   VAR CONSTANT
      C_REF_FREQUENCY : Int := 6000;   // [rpm]
      C_REF_VOLTAGE : Int := 1000;   // [V]
      C_REF_CURRENT : Int := 10;   // [A]
      C_REF_TORQUE : Int := 100;   // [Nm]
      C_REF_POWER : Int := 31;   // [W]
      C_REF_TEMP : Int := 100;   // [°C]
   END_VAR


BEGIN
	REGION Telegram Module
	    #t_ZSW1_Word := 0;
	    #t_POS_ZSW1_Word := 0;
	    #t_POS_ZSW2_Word := 0;
	    #t_ZSW2_Word := 0;

	    #t_Ret_Val_Int := RD_ADDR(LADDR := #i_Telegram_HW_ID,
	                              PIADDR => #t_HW_RD_Inf_Rec_I_Address,
	                              PICount => #t_HW_RD_Inf_Rec_I_Len,
	                              PQADDR => #t_HW_WR_Inf_Rec_O_Address,
	                              PQCount => #t_HW_WR_Inf_Rec_O_Len);

	    #o_Telegram_Start_Address := UDINT_TO_INT(#t_HW_RD_Inf_Rec_I_Address);

	    IF #t_Ret_Val_Int = 0 AND #t_HW_RD_Inf_Rec_I_Len = 24 THEN
	        // PZD1: ZSW1 (Word)
	        #t_ZSW1_Word := PEEK_WORD(area := 16#81, // Input area
	                                  dbNumber := 0,
	                                  byteOffset := UDINT_TO_DINT(#t_HW_RD_Inf_Rec_I_Address));

	        // PZD2: POS_ZSW1 (Word)
	        #t_POS_ZSW1_Word := PEEK_WORD(area := 16#81,
	                                      dbNumber := 0,
	                                      byteOffset := UDINT_TO_DINT(#t_HW_RD_Inf_Rec_I_Address) + 2);

	        // PZD3: POS_ZSW2 (Word)
	        #t_POS_ZSW2_Word := PEEK_WORD(area := 16#81,
	                                      dbNumber := 0,
	                                      byteOffset := UDINT_TO_DINT(#t_HW_RD_Inf_Rec_I_Address) + 4);

	        // PZD4: ZSW2 (Word)
	        #t_ZSW2_Word := PEEK_WORD(area := 16#81,
	                                  dbNumber := 0,
	                                  byteOffset := UDINT_TO_DINT(#t_HW_RD_Inf_Rec_I_Address) + 6);

	        // PZD5: Reserved (Int)
	        #o_Data.Reserved := 0;

	        // PZD6-7: XIST (Real/Float32) - Position actual value
	        #o_Data.XIST := DWORD_TO_REAL(PEEK_DWORD(area := 16#81,
	                                                                               dbNumber := 0,
	                                                                               byteOffset := UDINT_TO_DINT(#t_HW_RD_Inf_Rec_I_Address) + 10));

	        // PZD8-9: VIST (Real/Float32) - Velocity actual value
	        #o_Data.VIST := DWORD_TO_REAL(PEEK_DWORD(area := 16#81,
	                                                                               dbNumber := 0,
	                                                                               byteOffset := UDINT_TO_DINT(#t_HW_RD_Inf_Rec_I_Address) + 14));

	        // PZD10: MELDW (Word)
	        #o_Data.MELDW_Bit00_PositioningAbsolute := FALSE; // MELDW reserved in telegram 112

	        // PZD11: FaultCode (Word)
	        #o_Data.FaultCode := PEEK_WORD(area := 16#81,
	                                       dbNumber := 0,
	                                       byteOffset := UDINT_TO_DINT(#t_HW_RD_Inf_Rec_I_Address) + 20);

	        // PZD12: AlarmCode (Word)
	        #o_Data.AlarmCode := PEEK_WORD(area := 16#81,
	                                      dbNumber := 0,
	                                      byteOffset := UDINT_TO_DINT(#t_HW_RD_Inf_Rec_I_Address) + 22);
	    ELSE
	        #o_Data.XIST := 0.0;
	        #o_Data.VIST := 0.0;
	        #o_Data.FaultCode := 0;
	        #o_Data.AlarmCode := 0;
	    END_IF;

	    // Unpack ZSW1 bits
	    #o_Data.ZSW1_Bit00_ReadyOn := #t_ZSW1_Word.%X0;
	    #o_Data.ZSW1_Bit01_Ready := #t_ZSW1_Word.%X1;
	    #o_Data.ZSW1_Bit02_Enabled := #t_ZSW1_Word.%X2;
	    #o_Data.ZSW1_Bit03_Fault := #t_ZSW1_Word.%X3;
	    #o_Data.ZSW1_Bit04_Off2Inactive := #t_ZSW1_Word.%X4;
	    #o_Data.ZSW1_Bit05_Off3Inactive := #t_ZSW1_Word.%X5;
	    #o_Data.ZSW1_Bit06_Inhibit := #t_ZSW1_Word.%X6;
	    #o_Data.ZSW1_Bit07_Alarm := #t_ZSW1_Word.%X7;
	    #o_Data.ZSW1_Bit08_FollowingOK := #t_ZSW1_Word.%X8;
	    #o_Data.ZSW1_Bit09_Control := #t_ZSW1_Word.%X9;
	    #o_Data.ZSW1_Bit10_TargetReached := #t_ZSW1_Word.%X10;
	    #o_Data.ZSW1_Bit11_HomeSet := #t_ZSW1_Word.%X11;
	    #o_Data.ZSW1_Bit12_AckActive := #t_ZSW1_Word.%X12;
	    #o_Data.ZSW1_Bit13_SetpointFixed := #t_ZSW1_Word.%X13;
	    #o_Data.ZSW1_Bit14_AxisAccel := #t_ZSW1_Word.%X14;
	    #o_Data.ZSW1_Bit15_AxisDecel := #t_ZSW1_Word.%X15;

	    // Unpack POS_ZSW1 bits
	    #o_Data.POS_ZSW1_Bit00_Active0 := #t_POS_ZSW1_Word.%X0;
	    #o_Data.POS_ZSW1_Bit01_Active1 := #t_POS_ZSW1_Word.%X1;
	    #o_Data.POS_ZSW1_Bit02_Active2 := #t_POS_ZSW1_Word.%X2;
	    #o_Data.POS_ZSW1_Bit03_Active3 := #t_POS_ZSW1_Word.%X3;
	    #o_Data.POS_ZSW1_Bit04_Active4 := #t_POS_ZSW1_Word.%X4;
	    #o_Data.POS_ZSW1_Bit05_Active5 := #t_POS_ZSW1_Word.%X5;
	    #o_Data.POS_ZSW1_Bit06_Reserved := #t_POS_ZSW1_Word.%X6;
	    #o_Data.POS_ZSW1_Bit07_ReleaseBrake := #t_POS_ZSW1_Word.%X7;
	    #o_Data.POS_ZSW1_Bit08_StopCamMinus := #t_POS_ZSW1_Word.%X8;
	    #o_Data.POS_ZSW1_Bit09_StopCamPlus := #t_POS_ZSW1_Word.%X9;
	    #o_Data.POS_ZSW1_Bit10_JogActive := #t_POS_ZSW1_Word.%X10;
	    #o_Data.POS_ZSW1_Bit11_RefApproach := #t_POS_ZSW1_Word.%X11;
	    #o_Data.POS_ZSW1_Bit12_FlyingHoming := #t_POS_ZSW1_Word.%X12;
	    #o_Data.POS_ZSW1_Bit13_Traversing := #t_POS_ZSW1_Word.%X13;
	    #o_Data.POS_ZSW1_Bit14_Setup := #t_POS_ZSW1_Word.%X14;
	    #o_Data.POS_ZSW1_Bit15_MDI := #t_POS_ZSW1_Word.%X15;

	    // Unpack POS_ZSW2 bits
	    #o_Data.POS_ZSW2_Bit00_Tracking := #t_POS_ZSW2_Word.%X0;
	    #o_Data.POS_ZSW2_Bit01_VelLimit := #t_POS_ZSW2_Word.%X1;
	    #o_Data.POS_ZSW2_Bit02_TargetReached := #t_POS_ZSW2_Word.%X2;
	    #o_Data.POS_ZSW2_Bit03_PrintMark := #t_POS_ZSW2_Word.%X3;
	    #o_Data.POS_ZSW2_Bit04_Forward := #t_POS_ZSW2_Word.%X4;
	    #o_Data.POS_ZSW2_Bit05_Backward := #t_POS_ZSW2_Word.%X5;
	    #o_Data.POS_ZSW2_Bit06_SWLimitMinus := #t_POS_ZSW2_Word.%X6;
	    #o_Data.POS_ZSW2_Bit07_SWLimitPlus := #t_POS_ZSW2_Word.%X7;
	    #o_Data.POS_ZSW2_Bit08_Cam1 := #t_POS_ZSW2_Word.%X8;
	    #o_Data.POS_ZSW2_Bit09_Cam2 := #t_POS_ZSW2_Word.%X9;
	    #o_Data.POS_ZSW2_Bit10_Output1 := #t_POS_ZSW2_Word.%X10;
	    #o_Data.POS_ZSW2_Bit11_Output2 := #t_POS_ZSW2_Word.%X11;
	    #o_Data.POS_ZSW2_Bit12_FixedStop := #t_POS_ZSW2_Word.%X12;
	    #o_Data.POS_ZSW2_Bit13_Clamping := #t_POS_ZSW2_Word.%X13;
	    #o_Data.POS_ZSW2_Bit14_TravelFixed := #t_POS_ZSW2_Word.%X14;
	    #o_Data.POS_ZSW2_Bit15_TraversingCmd := #t_POS_ZSW2_Word.%X15;

	    // Unpack ZSW2 bits
	    #o_Data.ZSW2_Bit00_Reserved := #t_ZSW2_Word.%X0;
	    #o_Data.ZSW2_Bit01_Reserved := #t_ZSW2_Word.%X1;
	    #o_Data.ZSW2_Bit02_Reserved := #t_ZSW2_Word.%X2;
	    #o_Data.ZSW2_Bit03_Reserved := #t_ZSW2_Word.%X3;
	    #o_Data.ZSW2_Bit04_Reserved := #t_ZSW2_Word.%X4;
	    #o_Data.ZSW2_Bit05_Reserved := #t_ZSW2_Word.%X5;
	    #o_Data.ZSW2_Bit06_Reserved := #t_ZSW2_Word.%X6;
	    #o_Data.ZSW2_Bit07_Reserved := #t_ZSW2_Word.%X7;
	    #o_Data.ZSW2_Bit08_Reserved := #t_ZSW2_Word.%X8;
	    #o_Data.ZSW2_Bit09_Reserved := #t_ZSW2_Word.%X9;
	    #o_Data.ZSW2_Bit10_Reserved := #t_ZSW2_Word.%X10;
	    #o_Data.ZSW2_Bit11_Reserved := #t_ZSW2_Word.%X11;
	    #o_Data.ZSW2_Bit12_Reserved := #t_ZSW2_Word.%X12;
	    #o_Data.ZSW2_Bit13_Reserved := #t_ZSW2_Word.%X13;
	    #o_Data.ZSW2_Bit14_Reserved := #t_ZSW2_Word.%X14;
	    #o_Data.ZSW2_Bit15_Reserved := #t_ZSW2_Word.%X15;
	END_REGION

	REGION Actual Value Module (Extended Data)
	    #t_ZSW_S210_Word := 0;

	    #t_Ret_Val_Int := RD_ADDR(LADDR := #i_Additional_HW_ID,
	                              PIADDR => #t_HW_RD_Inf_Rec_I_Address,
	                              PICount => #t_HW_RD_Inf_Rec_I_Len,
	                              PQADDR => #t_HW_WR_Inf_Rec_O_Address,
	                              PQCount => #t_HW_WR_Inf_Rec_O_Len);

	    #o_ActualValue_Start_Address := UDINT_TO_INT(#t_HW_RD_Inf_Rec_I_Address);

	    IF #t_Ret_Val_Int = 0 AND #t_HW_RD_Inf_Rec_I_Len = 12 THEN
	        // Read ZSW_S210 (DI status word)
	        #t_ZSW_S210_Word := PEEK_WORD(area := 16#81, // Input area
	                                      dbNumber := 0,
	                                      byteOffset := UDINT_TO_DINT(#t_HW_RD_Inf_Rec_I_Address));

	        // Read DC Link Voltage (Int)
	        #t_Word_Scale_Data := PEEK_WORD(area := 16#81,
	                                        dbNumber := 0,
	                                        byteOffset := UDINT_TO_DINT(#t_HW_RD_Inf_Rec_I_Address) + 2);

	        #o_Data.DCLinkVoltage := DINT_TO_INT(WORD_TO_DINT(#t_Word_Scale_Data) * #C_REF_VOLTAGE / 16#4000);

	        // Read Actual Current (Int)
	        #t_Word_Scale_Data := PEEK_WORD(area := 16#81,
	                                        dbNumber := 0,
	                                        byteOffset := UDINT_TO_DINT(#t_HW_RD_Inf_Rec_I_Address) + 4);

	        #o_Data.ActualCurrent := DINT_TO_INT(WORD_TO_DINT(#t_Word_Scale_Data) * #C_REF_CURRENT * 10 / 16#4000);

	        // Read Active Power (Int)
	        #t_Word_Scale_Data := PEEK_WORD(area := 16#81,
	                                        dbNumber := 0,
	                                        byteOffset := UDINT_TO_DINT(#t_HW_RD_Inf_Rec_I_Address) + 6);

	        #o_Data.ActivePower := DINT_TO_INT(WORD_TO_DINT(#t_Word_Scale_Data) * #C_REF_POWER / 16#4000);

	        // Read Active Utilization (Int)
	        #t_Word_Scale_Data := PEEK_WORD(area := 16#81,
	                                        dbNumber := 0,
	                                        byteOffset := UDINT_TO_DINT(#t_HW_RD_Inf_Rec_I_Address) + 8);

	        #o_Data.TorqueUtilization := DINT_TO_INT(WORD_TO_DINT(#t_Word_Scale_Data) * 100 / 16#4000);

	        // Read Motor Load Rate (Int)
	        #t_Word_Scale_Data := PEEK_WORD(area := 16#81,
	                                        dbNumber := 0,
	                                        byteOffset := UDINT_TO_DINT(#t_HW_RD_Inf_Rec_I_Address) + 10);

	        #o_Data.MotorUtilization := DINT_TO_INT(WORD_TO_DINT(#t_Word_Scale_Data) * 100 / 16#4000);
	    ELSE
	        #o_Data.DCLinkVoltage := 0;
	        #o_Data.ActualCurrent := 0;
	        #o_Data.ActivePower := 0;
	        #o_Data.TorqueUtilization := 0;
	        #o_Data.MotorUtilization := 0;
	    END_IF;

	    // Unpack ZSW_S210 bits (DI status)
	    #o_Data.ZSW_S210_Bit00_DI0 := #t_ZSW_S210_Word.%X0;
	    #o_Data.ZSW_S210_Bit01_DI1 := #t_ZSW_S210_Word.%X1;
	    #o_Data.ZSW_S210_Bit02_DI2 := #t_ZSW_S210_Word.%X2;
	    #o_Data.ZSW_S210_Bit03_DI3 := #t_ZSW_S210_Word.%X3;
	    #o_Data.ZSW_S210_Bit04_DI4 := #t_ZSW_S210_Word.%X4;
	    #o_Data.ZSW_S210_Bit05_Reserved := #t_ZSW_S210_Word.%X5;
	    #o_Data.ZSW_S210_Bit06_Reserved := #t_ZSW_S210_Word.%X6;
	    #o_Data.ZSW_S210_Bit07_Reserved := #t_ZSW_S210_Word.%X7;
	    #o_Data.ZSW_S210_Bit08_Reserved := #t_ZSW_S210_Word.%X8;
	    #o_Data.ZSW_S210_Bit09_Reserved := #t_ZSW_S210_Word.%X9;
	    #o_Data.ZSW_S210_Bit10_Reserved := #t_ZSW_S210_Word.%X10;
	    #o_Data.ZSW_S210_Bit11_Reserved := #t_ZSW_S210_Word.%X11;
	    #o_Data.ZSW_S210_Bit12_Reserved := #t_ZSW_S210_Word.%X12;
	    #o_Data.ZSW_S210_Bit13_Reserved := #t_ZSW_S210_Word.%X13;
	    #o_Data.ZSW_S210_Bit14_Reserved := #t_ZSW_S210_Word.%X14;
	    #o_Data.ZSW_S210_Bit15_Reserved := #t_ZSW_S210_Word.%X15;
	END_REGION
END_FUNCTION

TYPE "UDT_S210_SW_Output"
VERSION : 0.1
   STRUCT
      AxisEnabled : Bool;   // 驱动已使能
      AxisPosOk : Bool;   // 目标位置到达
      AxisSpFixed : Bool;   // 设定位置到达
      AxisRef : Bool;   // 已设置参考点
      AxisWarn : Bool;   // 驱动报警
      AxisError : Bool;   // 驱动故障
      Lockout : Bool;   // 禁止接通
      ActVelocity : Real;   // 实际速度
      ActPosition : Real;   // 当前位置
      ActMode : Int;   // 当前激活的运行模式
      EPosZSW1 : Word;   // POS ZSW1的状态
      EPosZSW2 : Word;   // POS ZSW2的状态
      AlarmCode : Word;   // 驱动器当前的报警代码
      FaultCode : Word;   // 驱动器当前的故障代码
      ZSW1 : Word;   // ZSW1的状态
      ZSW2 : Word;   // ZSW2的状态
      MELDW : Word;   // MELDW的状态
      Error : Bool;   // 1=存在错误
      Status : Word;   // 16#7002：无故障，正常运行
      DiagID : Word;   // 扩展的通信错误
   END_STRUCT;

END_TYPE

TYPE "UDT_S210_SW_Input"
VERSION : 0.1
   STRUCT
      Mode : Int;
      Enbale : Bool;
      CancelTraversing : Bool;
      IntermediateStop : Bool;
      Positive : Bool;
      Negative : Bool;
      Jog_Left : Bool;
      Jog_Right : Bool;
      FlyRef : Bool;
      AckError : Bool;
      ExecuteMode : Bool;
      Position : Real;
      Velocity : Real;
      OverV : Int;
      Acceleration : Real;
      Deceleration : Real;
      FixStopTorque : Real;
      RefCoordinate : Real;
      ConfigEPOS : DWord;
   END_STRUCT;

END_TYPE

FUNCTION_BLOCK "FB_SINA_POS_TEL112"
{ S7_Optimized_Access := 'TRUE' }
VERSION : 0.2
   VAR_INPUT
      modePos : Int;   // Settings of the mode
      enableAxis : Bool;   // 1 = Enable the drive
      cancelTraversing : Bool := TRUE;   // 0 = Reject active traverse task
      intermediateStop : Bool := TRUE;   // 0 = Intermediate STOP of traverse command
      positive : Bool;   // 1 = Direction positive
      negative : Bool;   // 1 = Direction negative
      jog1 : Bool;   // 1 = Use jog 1 (direction / speed)
      jog2 : Bool;   // 1 = Use jog 2 (direction / speed)
      flyRef : Bool;   // 1 = Start flying reference function
      ackError : Bool;   // 1  = Acknowledge of errors
      executeMode : Bool;   // 0-->1 = Start the mode
      position : Real;   // Position of the MDI mode or setting of traversing block
      velocity : Real;   // MDI velocity
      overV : Int := 100;   // Override of  velocity in [%] --> 4000h=100%
      acceleration : Real;   // MDI acceleration
      deceleration : Real;   // MDI deceleration
      fixStopTorque : Real;   // torque setting for fix stop function (reserved)
      refCoordinate : Real;
      configEPOS : DWord := 16#0000_0003;   // binary programmed input to control all functions in the telegram without its own function block input
   END_VAR

   VAR_OUTPUT
      axisEnabled : Bool;   // 1= Axis in operation
      axisPosOk : Bool;   // 1= Position setpoint reached
      axisSpFixed : Bool;   // 1= Setpoint fixed (Attention: Dependence on SINAMICS firmware)
      axisRef : Bool;   // 1= Reference point set
      axisWarn : Bool;   // 1= Axis alarm / warning present
      axisError : Bool;   // 1= Axis fault present
      lockOut : Bool;   // 1= Axis in lockout state
      actVelocity : Real;   // actual axis velocity
      actPosition : Real;   // actual axis position
      actMode : Int;   // Active EPos mode
      actWarn : Word;   // Actual number of warning
      actFault : Word;   // Actual number of error
      error : Bool;   // 1 = Error  (FB and Infeed)
      status : Word;   // Status output (7002 = FB in operation; 8xxx = error description  - read the manual)
      diagID : Word;   // Error codes of the cyclic system funtion blocks DPWR / DPRD_DAT (固定为0)
   END_VAR

   VAR_IN_OUT
      InputData : "UDT_S210_HW_Input";   // 从驱动器接收的数据
      OutputData : "UDT_S210_HW_Output";   // 发送到驱动器的数据
   END_VAR

   VAR
      sbOff1Edge : Bool := 0;   // Positive edge of starting or stopping the device
      sbOff1 : Bool := 0;   // Starting or stopping the device
      sbExecuteEdge : Bool := 0;   // Positive edge of activate traversing block
      sbExecute : Bool := 0;   // Activate traversing block
      sbRefTypEdge : Bool := 0;   // Positive edge of referencing type "flying reference"
      sbRefTyp : Bool := 0;   // Referencing type "flying reference"
      sbMdiStart : Bool := 0;   // Direct setpoint input / MDI - start
      sbMdiStartEdge : Bool := 0;   // Positive edge of direct setpoint input / MDI - start
      sbRefStart : Bool := 0;   // Referencing start
      sbJogInc : Bool := 0;   // Jogging incremental
      sbReady : Bool := 0;   // Ready to power up / to start
      sbIOp : Bool := 0;   // Ready to operate
      sbAccel : Bool := 0;   // Axis accelerating
      sbDecel : Bool := 0;   // Axis decelerating
      sbAlarm : Bool := 0;   // Alarm / Warnung present
      sbFault : Bool := 0;   // Fault present
      sbFWD : Bool := 0;   // Axis drives forwards
      sbBWD : Bool := 0;   // Axis drives backwards
      sbBusy : Bool := 0;   // Mode of operation is explained
      swStatus : Word := 16#0000;   // Mode of operation disturbance
      siExecuteCyc : Int := 0;   // Counter of runcycle of active traversing block
      siRefTypCyc : Int := 0;   // Counter of runcycle of referencing type "flying reference"
      siJogIncCyc : Int := 0;   // Counter of runcycle of jogging incremental
      siMdiStartCyc : Int := 0;   // Counter of runcycle of direct setpoint input / MDI - start
      siRefActRetry : Int := 0;   // Counter of retry of reference point approach active
      siModePos : Int := 0;   // Setting of mode
      siCycWait : Int := 5;   // Counter of cycle of waiting
      siRetryMax : Int := 30;   // Max. count of cycles of retry
      sbModePos : Bool := 0;   // Mode of setting okay
   END_VAR

   VAR CONSTANT
      MODEPOSMAX : Int := 9;   // Max. count of mode
      TRAVERSEBLOCKMAXNO : Int := 32;   // Max. number of traversing block
   END_VAR


BEGIN
	//=============================================================================
	//SIEMENS AG
	//(c)Copyright 2023 All Rights Reserved
	//-----------------------------------------------------------------------------
	// Library: DriveLib
	// Tested with: -
	// Engineering: TIA Portal V18
	// Restrictions: -
	// Requirements: S7-1200 / S7-1500
	// Functionality: cyclic communication between a SINAMICS (Basic positioner)and a PLC
	//                If in HWConfig Std.TLG 112 is projected 17/12 PZD-words are exchanged
	//                in every bus cycle.
	//                The parametrisation of these words is described in the manual of the
	//                SINAMICS
	// Contactor: mc_gmc_mp_asia.cn@siemens.com
	// *****************************************************************************
	// Version:
	// V0.0: Created
	// V0.2: 重构 - 移除DPWR/DPRD，改用外部UDT (UDT_S210_HW_Output/Input)
	//=============================================================================

	// The input of the modePos should between 1 and the MODEPOSMAX
	IF #modePos > #MODEPOSMAX OR #modePos < 1 THEN
	    #sbModePos := FALSE;
	    #error := True;
	    #swStatus := 16#8202;
	ELSE
	    IF NOT #sbFWD AND NOT #sbBWD AND NOT #sbAccel AND NOT #sbDecel THEN
	        #sbModePos := TRUE;
	        #siModePos := #modePos;
	        IF #swStatus = 16#8202 THEN
	            #swStatus := 16#7002;
	            #error := False;
	        END_IF;
	    END_IF;
	END_IF;

	// Check the overrider setting
	IF (#overV < 0) OR (#overV > 199) THEN
	    #swStatus := 16#8203;
	    #error := True;
	ELSE
	    // Override映射到OutputData.Override (Int类型，0-16384对应0-100%)
	    #OutputData.Override := REAL_TO_INT(16384.0 * (INT_TO_REAL(#overV) / 100.0));
	END_IF;

	// Check the acceleration and deceleration setting
	IF #acceleration < 0.0 THEN
	    #swStatus := 16#8203;
	    #error := True;
	ELSE
	    #OutputData.MDI_ACC := #acceleration;
	END_IF;
	IF #deceleration < 0.0 THEN
	    #swStatus := 16#8203;
	    #error := True;
	ELSE
	    #OutputData.MDI_DEC := #deceleration;
	END_IF;
	IF NOT (#overV < 0) AND NOT (#overV > 199) AND NOT (#acceleration < 0.0) AND NOT (#deceleration < 0.0) THEN
	    IF #swStatus = 16#8203 THEN
	        #swStatus := 16#7002;
	        #error := FALSE;
	    END_IF;
	END_IF;

	// 位置、速度、参考坐标直接映射
	#OutputData.MDI_TARPOS := #position;
	#OutputData.MDI_VELOCITY := #velocity;
	#OutputData.REF_COORDINATE := #refCoordinate;

	// Enable the axis
	IF #enableAxis AND NOT #sbOff1Edge AND NOT #sbBusy AND #sbModePos THEN
	    #sbOff1 := True;
	END_IF;
	#sbOff1Edge := #enableAxis AND NOT #sbBusy;
	IF NOT #enableAxis THEN
	    #sbOff1 := False;
	END_IF;

	// Flying reference
	IF #flyRef AND NOT #sbRefTypEdge THEN
	    #sbRefTyp := True;
	END_IF;
	#sbRefTypEdge := #flyRef;
	IF NOT #flyRef THEN
	    #sbRefTyp := False;
	    #siRefTypCyc := 0;
	END_IF;

	// Execute the motion
	IF #executeMode AND NOT #sbExecuteEdge THEN
	    #sbExecute := True;
	    #siExecuteCyc := 0;
	ELSIF #actMode <> #modePos THEN
	    #sbExecute := FALSE;
	ELSIF #siExecuteCyc > (15 * #siCycWait) THEN
	    IF #modePos <> 4 THEN
	        #sbExecute := FALSE;
	    ELSE
	        // 使用InputData.ZSW1_Bit11_HomeSet替代sxRecvBuf.ZSW1.%X11
	        IF #InputData.ZSW1_Bit11_HomeSet OR NOT #executeMode THEN
	            #sbExecute := FALSE;
	        END_IF;
	    END_IF;
	ELSE
	    ;
	END_IF;
	IF #siExecuteCyc > 100 THEN
	    #siExecuteCyc := 0;
	ELSE
	    #siExecuteCyc := #siExecuteCyc + 1;
	END_IF;
	#sbExecuteEdge := #executeMode;

	// MDI Start边沿检测逻辑（基于EPosSTW1.%X15，即POS_STW1_Bit15_ActivateMDI）
	IF #OutputData.POS_STW1_Bit15_ActivateMDI AND NOT #sbMdiStartEdge THEN
	    #sbMdiStart := True;
	END_IF;
	#sbMdiStartEdge := #OutputData.POS_STW1_Bit15_ActivateMDI AND NOT #sbBusy;
	IF NOT #OutputData.POS_STW1_Bit15_ActivateMDI THEN
	    #sbMdiStart := False;
	    #siMdiStartCyc := 0;
	END_IF;

	// 基础STW1控制位映射
	#OutputData.STW1_Bit04_NotRejectTask := #cancelTraversing;
	#OutputData.STW1_Bit05_NoIntermediateStop := #intermediateStop;
	#OutputData.STW1_Bit07_Ack := #ackError;
	#OutputData.STW1_Bit01_Off2 := TRUE;  // 原.%X1
	#OutputData.STW1_Bit02_Off3 := TRUE;  // 原.%X2
	#OutputData.STW1_Bit03_Enable := TRUE; // 原.%X3
	#OutputData.STW1_Bit10_PLC := TRUE;    // 原.%X10 (Life bit)
	#OutputData.STW1_Bit12_Reserved := FALSE; // 原.%X12
	#OutputData.STW1_Bit14_Reserved := FALSE; // 原.%X14
	#OutputData.STW1_Bit15_Reserved := FALSE; // 原.%X15

	// If the parameter setting is correnct, then execute the positioning mode.
	// ModePos = 1, relative positioning
	IF (#siModePos = 1 AND #sbModePos) THEN
	    #OutputData.STW1_Bit00_On := #sbOff1;           // 原STW1.%X0
	    #OutputData.STW1_Bit08_Jog1 := False;           // 原.%X8
	    #OutputData.STW1_Bit09_Jog2 := False;           // 原.%X9
	    #OutputData.STW1_Bit11_StartHoming := False;    // 原.%X11

	    #OutputData.POS_STW1_Bit08_Absolute := False;    // 原EPosSTW1.%X8 (0=相对)
	    #OutputData.POS_STW1_Bit09_DirPos := False;      // 原.%X9
	    #OutputData.POS_STW1_Bit10_DirNeg := False;      // 原.%X10
	    #OutputData.POS_STW1_Bit14_SetupOrPositioning := False; // 原.%X14 (0=定位)
	    #OutputData.POS_STW1_Bit15_ActivateMDI := False; // 原.%X15

	    #OutputData.POS_STW2_Bit01_SetRefPoint := False;  // 原.%X1
	    #OutputData.POS_STW2_Bit03_AdjustEncoder := False; // 原.%X3
	    #OutputData.POS_STW2_Bit05_JogIncrementalOrVelocity := False; // 原.%X5
	    #OutputData.POS_STW2_Bit09_RefNegDir := False;    // 原.%X9
	    #OutputData.POS_STW2_Bit08_RefType := False;      // 原.%X8

	    IF #sbOff1 AND #sbReady AND #sbIOp AND NOT #sbFault THEN
	        #OutputData.POS_STW1_Bit15_ActivateMDI := True;  // MDI激活
	        #OutputData.POS_STW1_Bit08_Absolute := False;    // 相对定位
	        IF #positive AND NOT #negative THEN
	            #OutputData.POS_STW1_Bit09_DirPos := True;
	            #OutputData.POS_STW1_Bit10_DirNeg := False;
	        ELSIF NOT #positive AND #negative THEN
	            #OutputData.POS_STW1_Bit09_DirPos := False;
	            #OutputData.POS_STW1_Bit10_DirNeg := True;
	        ELSE
	            #OutputData.POS_STW1_Bit09_DirPos := False;
	            #OutputData.POS_STW1_Bit10_DirNeg := False;
	        END_IF;
	        IF #sbMdiStart AND (#siMdiStartCyc < #siCycWait) THEN
	            #siMdiStartCyc := #siMdiStartCyc + 1;
	        ELSE
	            #OutputData.STW1_Bit06_ActivateTask := #sbExecute; // 原.%X6
	        END_IF;
	        IF #sbRefTyp THEN
	            #OutputData.POS_STW2_Bit08_RefType := True; // 飞参模式
	            IF (#siRefTypCyc = 0) THEN
	                #siRefTypCyc := #siRefTypCyc + 1;
	            ELSE
	                #OutputData.STW1_Bit11_StartHoming := True; // 开始回零
	            END_IF;
	        END_IF;
	    END_IF;

	    // ModePos = 2, absolute positioning
	ELSIF (#siModePos = 2 AND #sbModePos) THEN
	    #OutputData.STW1_Bit00_On := #sbOff1;
	    #OutputData.STW1_Bit08_Jog1 := False;
	    #OutputData.STW1_Bit09_Jog2 := False;
	    #OutputData.STW1_Bit11_StartHoming := False;

	    #OutputData.POS_STW1_Bit08_Absolute := False;
	    #OutputData.POS_STW1_Bit09_DirPos := False;
	    #OutputData.POS_STW1_Bit10_DirNeg := False;
	    #OutputData.POS_STW1_Bit14_SetupOrPositioning := False;
	    #OutputData.POS_STW1_Bit15_ActivateMDI := False;

	    #OutputData.POS_STW2_Bit01_SetRefPoint := False;
	    #OutputData.POS_STW2_Bit03_AdjustEncoder := False;
	    #OutputData.POS_STW2_Bit05_JogIncrementalOrVelocity := False;
	    #OutputData.POS_STW2_Bit09_RefNegDir := False;
	    #OutputData.POS_STW2_Bit08_RefType := False;

	    IF #sbOff1 AND #sbReady AND #sbIOp AND NOT #sbFault THEN
	        #OutputData.POS_STW1_Bit15_ActivateMDI := True;
	        #OutputData.POS_STW1_Bit08_Absolute := True;  // 绝对定位
	        IF #positive AND NOT #negative THEN
	            #OutputData.POS_STW1_Bit09_DirPos := True;
	            #OutputData.POS_STW1_Bit10_DirNeg := False;
	        ELSIF NOT #positive AND #negative THEN
	            #OutputData.POS_STW1_Bit09_DirPos := False;
	            #OutputData.POS_STW1_Bit10_DirNeg := True;
	        ELSE
	            #OutputData.POS_STW1_Bit09_DirPos := False;
	            #OutputData.POS_STW1_Bit10_DirNeg := False;
	        END_IF;
	        IF #sbMdiStart AND (#siMdiStartCyc < #siCycWait) THEN
	            #siMdiStartCyc := #siMdiStartCyc + 1;
	        ELSE
	            #OutputData.STW1_Bit06_ActivateTask := #sbExecute;
	        END_IF;
	        IF #sbRefTyp THEN
	            #OutputData.POS_STW2_Bit08_RefType := True;
	            IF (#siRefTypCyc = 0) THEN
	                #siRefTypCyc := #siRefTypCyc + 1;
	            ELSE
	                #OutputData.STW1_Bit11_StartHoming := True;
	            END_IF;
	        END_IF;
	    END_IF;

	    // ModePos = 3, setup mode
	ELSIF (#siModePos = 3 AND #sbModePos) THEN
	    #OutputData.STW1_Bit00_On := #sbOff1;
	    #OutputData.STW1_Bit08_Jog1 := False;
	    #OutputData.STW1_Bit09_Jog2 := False;
	    #OutputData.STW1_Bit11_StartHoming := False;

	    #OutputData.POS_STW1_Bit08_Absolute := False;
	    #OutputData.POS_STW1_Bit09_DirPos := False;
	    #OutputData.POS_STW1_Bit10_DirNeg := False;
	    #OutputData.POS_STW1_Bit14_SetupOrPositioning := False;
	    #OutputData.POS_STW1_Bit15_ActivateMDI := False;

	    #OutputData.POS_STW2_Bit01_SetRefPoint := False;
	    #OutputData.POS_STW2_Bit03_AdjustEncoder := False;
	    #OutputData.POS_STW2_Bit05_JogIncrementalOrVelocity := False;
	    #OutputData.POS_STW2_Bit09_RefNegDir := False;
	    #OutputData.POS_STW2_Bit08_RefType := False;

	    IF #sbOff1 AND #sbReady AND #sbIOp AND NOT #sbFault THEN
	        #OutputData.POS_STW1_Bit15_ActivateMDI := True;
	        #OutputData.POS_STW1_Bit08_Absolute := True;
	        #OutputData.POS_STW1_Bit14_SetupOrPositioning := True; // Setup模式
	        IF #positive AND NOT #negative THEN
	            #OutputData.POS_STW1_Bit09_DirPos := True;
	            #OutputData.POS_STW1_Bit10_DirNeg := False;
	        ELSIF NOT #positive AND #negative THEN
	            #OutputData.POS_STW1_Bit09_DirPos := False;
	            #OutputData.POS_STW1_Bit10_DirNeg := True;
	        ELSE
	            #OutputData.POS_STW1_Bit09_DirPos := False;
	            #OutputData.POS_STW1_Bit10_DirNeg := False;
	        END_IF;
	        IF #sbMdiStart AND (#siMdiStartCyc < #siCycWait) THEN
	            #siMdiStartCyc := #siMdiStartCyc + 1;
	        ELSE
	            #OutputData.STW1_Bit06_ActivateTask := #sbExecute;
	        END_IF;
	        IF #sbRefTyp THEN
	            #OutputData.POS_STW2_Bit08_RefType := True;
	            IF (#siRefTypCyc = 0) THEN
	                #siRefTypCyc := #siRefTypCyc + 1;
	            ELSE
	                #OutputData.STW1_Bit11_StartHoming := True;
	            END_IF;
	        END_IF;
	    END_IF;

	    // ModePos = 4, reference point approach
	ELSIF (#siModePos = 4 AND #sbModePos) THEN
	    #OutputData.STW1_Bit00_On := #sbOff1;
	    #OutputData.STW1_Bit08_Jog1 := False;
	    #OutputData.STW1_Bit09_Jog2 := False;
	    #OutputData.STW1_Bit11_StartHoming := False;

	    #OutputData.POS_STW1_Bit15_ActivateMDI := False;
	    #OutputData.POS_STW2_Bit01_SetRefPoint := False;
	    #OutputData.POS_STW2_Bit03_AdjustEncoder := False;
	    #OutputData.POS_STW2_Bit05_JogIncrementalOrVelocity := False;
	    #OutputData.POS_STW2_Bit08_RefType := False;
	    #OutputData.POS_STW2_Bit09_RefNegDir := False;

	    IF #sbOff1 AND #sbReady AND #sbIOp AND NOT #sbFault THEN
	        #OutputData.STW1_Bit11_StartHoming := #sbExecute;
	        IF #positive AND NOT #negative THEN
	            #OutputData.POS_STW2_Bit09_RefNegDir := False; // 正方向
	        ELSIF NOT #positive AND #negative THEN
	            #OutputData.POS_STW2_Bit09_RefNegDir := True;  // 负方向
	        END_IF;
	    END_IF;

	    // ModePos = 5, set reference point
	ELSIF (#siModePos = 5 AND #sbModePos) THEN
	    #OutputData.STW1_Bit08_Jog1 := False;
	    #OutputData.STW1_Bit09_Jog2 := False;
	    #OutputData.STW1_Bit11_StartHoming := False;
	    #OutputData.POS_STW1_Bit15_ActivateMDI := False;
	    #OutputData.POS_STW2_Bit03_AdjustEncoder := False;
	    #OutputData.POS_STW2_Bit05_JogIncrementalOrVelocity := False;
	    #OutputData.POS_STW2_Bit08_RefType := False;
	    #OutputData.POS_STW2_Bit09_RefNegDir := False;
	    #OutputData.POS_STW2_Bit01_SetRefPoint := False;

	    IF NOT #sbFault THEN
	        #OutputData.POS_STW2_Bit01_SetRefPoint := #sbExecute; // 设置参考点
	    END_IF;

	    // ModePos = 6, traversing block function
	ELSIF (#siModePos = 6 AND #sbModePos) THEN
	    #OutputData.STW1_Bit00_On := #sbOff1;
	    #OutputData.STW1_Bit08_Jog1 := False;
	    #OutputData.STW1_Bit09_Jog2 := False;
	    #OutputData.STW1_Bit11_StartHoming := False;

	    #OutputData.POS_STW1_Bit08_Absolute := False;
	    #OutputData.POS_STW1_Bit09_DirPos := False;
	    #OutputData.POS_STW1_Bit10_DirNeg := False;
	    #OutputData.POS_STW1_Bit14_SetupOrPositioning := False;
	    #OutputData.POS_STW1_Bit15_ActivateMDI := False;

	    #OutputData.POS_STW2_Bit01_SetRefPoint := False;
	    #OutputData.POS_STW2_Bit03_AdjustEncoder := False;
	    #OutputData.POS_STW2_Bit05_JogIncrementalOrVelocity := False;
	    #OutputData.POS_STW2_Bit09_RefNegDir := False;
	    #OutputData.POS_STW2_Bit08_RefType := False;

	    // 遍历块选择位清零
	    #OutputData.POS_STW1_Bit00_Traversing0 := False;
	    #OutputData.POS_STW1_Bit01_Traversing1 := False;
	    #OutputData.POS_STW1_Bit02_Traversing2 := False;
	    #OutputData.POS_STW1_Bit03_Traversing3 := False;
	    #OutputData.POS_STW1_Bit04_Traversing4 := False;
	    #OutputData.POS_STW1_Bit05_Traversing5 := False;

	    IF (DINT_TO_INT(TRUNC(#position)) < 0) OR (DINT_TO_INT(TRUNC(#position)) > #TRAVERSEBLOCKMAXNO) THEN
	        #swStatus := 16#8204;
	        #error := True;
	    ELSE
	        IF #swStatus = 16#8204 THEN
	            #swStatus := 16#7002;
	            #error := False;
	        END_IF;
	        // 遍历块位选择 (Bit0-5)
	        IF (INT_TO_WORD(DINT_TO_INT(TRUNC(#position))) AND W#16#01) = W#16#01 THEN
	            #OutputData.POS_STW1_Bit00_Traversing0 := True;
	        END_IF;
	        IF (INT_TO_WORD(DINT_TO_INT(TRUNC(#position))) AND W#16#02) = W#16#02 THEN
	            #OutputData.POS_STW1_Bit01_Traversing1 := True;
	        END_IF;
	        IF (INT_TO_WORD(DINT_TO_INT(TRUNC(#position))) AND W#16#04) = W#16#04 THEN
	            #OutputData.POS_STW1_Bit02_Traversing2 := True;
	        END_IF;
	        IF (INT_TO_WORD(DINT_TO_INT(TRUNC(#position))) AND W#16#08) = W#16#08 THEN
	            #OutputData.POS_STW1_Bit03_Traversing3 := True;
	        END_IF;
	        IF (INT_TO_WORD(DINT_TO_INT(TRUNC(#position))) AND W#16#10) = W#16#10 THEN
	            #OutputData.POS_STW1_Bit04_Traversing4 := True;
	        END_IF;
	        IF (INT_TO_WORD(DINT_TO_INT(TRUNC(#position))) AND W#16#20) = W#16#20 THEN
	            #OutputData.POS_STW1_Bit05_Traversing5 := True;
	        END_IF;

	        IF #sbOff1 AND #sbReady AND #sbIOp AND NOT #sbFault THEN
	            #OutputData.STW1_Bit06_ActivateTask := #sbExecute;
	            IF #sbRefTyp THEN
	                #OutputData.POS_STW2_Bit08_RefType := True;
	                IF (#siRefTypCyc = 0) THEN
	                    #siRefTypCyc := #siRefTypCyc + 1;
	                ELSE
	                    #OutputData.STW1_Bit11_StartHoming := True;
	                END_IF;
	            END_IF;
	        END_IF;
	    END_IF;

	    // ModePos = 7, jog
	ELSIF (#siModePos = 7 AND #sbModePos) THEN
	    #OutputData.STW1_Bit00_On := #sbOff1;
	    #OutputData.STW1_Bit08_Jog1 := False;
	    #OutputData.STW1_Bit09_Jog2 := False;
	    #OutputData.STW1_Bit11_StartHoming := False;

	    #OutputData.POS_STW1_Bit15_ActivateMDI := False;
	    #OutputData.POS_STW2_Bit05_JogIncrementalOrVelocity := False;
	    #OutputData.POS_STW2_Bit08_RefType := False;
	    #OutputData.POS_STW2_Bit01_SetRefPoint := False;
	    #OutputData.POS_STW2_Bit03_AdjustEncoder := False;

	    IF #sbOff1 AND #sbReady AND #sbIOp AND NOT #sbFault THEN
	        IF #jog1 AND NOT #jog2 THEN
	            #OutputData.STW1_Bit08_Jog1 := True;
	        END_IF;
	        IF #jog2 AND NOT #jog1 THEN
	            #OutputData.STW1_Bit09_Jog2 := True;
	        END_IF;
	        IF #sbRefTyp THEN
	            #OutputData.POS_STW2_Bit08_RefType := #flyRef;
	            IF (#siRefTypCyc = 0) THEN
	                #siRefTypCyc := #siRefTypCyc + 1;
	            ELSE
	                #OutputData.STW1_Bit11_StartHoming := True;
	            END_IF;
	        END_IF;
	    END_IF;

	    // ModePos = 8, incremental jog
	ELSIF (#siModePos = 8 AND #sbModePos) THEN
	    #OutputData.STW1_Bit00_On := #sbOff1;
	    #OutputData.STW1_Bit08_Jog1 := False;
	    #OutputData.STW1_Bit09_Jog2 := False;
	    #OutputData.STW1_Bit11_StartHoming := False;

	    #OutputData.POS_STW1_Bit15_ActivateMDI := False;
	    #OutputData.POS_STW2_Bit05_JogIncrementalOrVelocity := False;
	    #OutputData.POS_STW2_Bit08_RefType := False;
	    #OutputData.POS_STW2_Bit01_SetRefPoint := False;
	    #OutputData.POS_STW2_Bit03_AdjustEncoder := False;

	    IF #sbOff1 AND #sbReady AND #sbIOp AND NOT #sbFault THEN
	        #OutputData.POS_STW2_Bit05_JogIncrementalOrVelocity := True; // 增量模式
	        #sbJogInc := True;
	        IF #sbJogInc AND (#siJogIncCyc = 0) THEN
	            #siJogIncCyc := #siJogIncCyc + 1;
	        ELSE
	            IF #jog1 XOR #jog2 THEN
	                #OutputData.STW1_Bit08_Jog1 := #jog1;
	                #OutputData.STW1_Bit09_Jog2 := #jog2;
	            END_IF;
	        END_IF;
	        IF #sbRefTyp THEN
	            #OutputData.POS_STW2_Bit08_RefType := True;
	            IF (#siRefTypCyc = 0) THEN
	                #siRefTypCyc := #siRefTypCyc + 1;
	            ELSE
	                #OutputData.STW1_Bit11_StartHoming := True;
	            END_IF;
	        END_IF;
	    END_IF;

	    // ModePos = 9 (Reserve/Encoder adjustment)
	ELSIF (#siModePos = 9 AND #sbModePos) THEN
	    #OutputData.STW1_Bit08_Jog1 := False;
	    #OutputData.STW1_Bit09_Jog2 := False;
	    #OutputData.STW1_Bit11_StartHoming := False;
	    #OutputData.POS_STW1_Bit15_ActivateMDI := False;
	    #OutputData.POS_STW2_Bit05_JogIncrementalOrVelocity := False;
	    #OutputData.POS_STW2_Bit08_RefType := False;
	    #OutputData.POS_STW2_Bit09_RefNegDir := False;
	    #OutputData.POS_STW2_Bit01_SetRefPoint := False;

	    IF NOT #sbFault THEN
	        #OutputData.POS_STW2_Bit03_AdjustEncoder := #sbExecute; // 编码器调整
	    END_IF;

	ELSE
	    // 默认状态/无效模式
	    #OutputData.STW1_Bit00_On := #enableAxis;
	    #OutputData.STW1_Bit04_NotRejectTask := False;
	    #OutputData.STW1_Bit06_ActivateTask := False;
	    #OutputData.POS_STW1_Bit15_ActivateMDI := False;
	    #OutputData.STW1_Bit08_Jog1 := False;
	    #OutputData.STW1_Bit09_Jog2 := False;
	    #OutputData.POS_STW1_Bit08_Absolute := False;
	    #OutputData.POS_STW1_Bit09_DirPos := False;
	    #OutputData.POS_STW1_Bit10_DirNeg := False;
	    #OutputData.POS_STW1_Bit12_Continuous := False;
	    #OutputData.POS_STW1_Bit14_SetupOrPositioning := False;
	    #OutputData.POS_STW2_Bit01_SetRefPoint := False;
	    #OutputData.POS_STW2_Bit08_RefType := False;
	    #OutputData.POS_STW2_Bit09_RefNegDir := False;
	    #OutputData.POS_STW2_Bit05_JogIncrementalOrVelocity := False;
	    #OutputData.POS_STW2_Bit03_AdjustEncoder := False;
	    #OutputData.STW1_Bit11_StartHoming := False;
	END_IF;

	// Configure the configEPOS to the telegram
	// 应用configEPOS映射（这些可能会覆盖上面的设置，根据原代码逻辑）
	#OutputData.STW1_Bit01_Off2 := #configEPOS.%X0;
	#OutputData.STW1_Bit02_Off3 := #configEPOS.%X1;
	#OutputData.STW1_Bit13_ExtBlockChange := #configEPOS.%X7;
	#OutputData.STW2_Bit08_Reserved := #configEPOS.%X30; // 注意：UDT中STW2保留，但原代码使用Bit8

	#OutputData.POS_STW1_Bit12_Continuous := #configEPOS.%X8;
	#OutputData.POS_STW2_Bit14_SWLimit := #configEPOS.%X2;
	#OutputData.POS_STW2_Bit15_StopCam := #configEPOS.%X3;
	#OutputData.POS_STW2_Bit11_MeasProbeEdge := #configEPOS.%X4;
	#OutputData.POS_STW2_Bit10_MeasProbe2 := #configEPOS.%X5;
	#OutputData.POS_STW2_Bit02_RefCam := #configEPOS.%X6;

	// 检查驱动器状态
	IF #InputData.ZSW1_Bit03_Fault THEN
	    #swStatus := 16#8401;
	    #error := True;
	ELSIF #InputData.ZSW1_Bit06_Inhibit THEN
	    #swStatus := 16#8402;
	    #error := True;
	ELSE
	    IF (#swStatus = 16#8401) OR (#swStatus = 16#8402) THEN
	        #swStatus := 16#7002;
	        #error := False;
	    END_IF;
	END_IF;

	// 飞参激活检测和重试逻辑（使用POS_ZSW1_Bit12_FlyingHoming）
	IF NOT #InputData.POS_ZSW1_Bit12_FlyingHoming AND #sbRefTyp AND #OutputData.STW1_Bit11_StartHoming THEN
	    IF #siRefActRetry < #siRetryMax THEN
	        #siRefActRetry := #siRefActRetry + 1;
	        #OutputData.STW1_Bit11_StartHoming := False;
	    ELSE
	        #swStatus := 16#8403;
	        #error := True;
	    END_IF;
	ELSE
	    IF #swStatus = 16#8403 THEN
	        #swStatus := 16#7002;
	        #error := False;
	    END_IF;
	    IF (#InputData.POS_ZSW1_Bit12_FlyingHoming AND #sbRefTyp AND #OutputData.STW1_Bit11_StartHoming) OR NOT #flyRef THEN
	        #siRefActRetry := 0;
	    END_IF;
	END_IF;

	// 诊断ID固定为0（无通信错误）
	#diagID := W#16#0000;

	// 处理接收数据 - 从InputData映射到内部变量和输出
	// 状态字ZSW1映射
	#sbReady := #InputData.ZSW1_Bit01_Ready;
	#axisEnabled := #InputData.ZSW1_Bit02_Enabled;
	#sbIOp := #InputData.ZSW1_Bit02_Enabled; // 同Bit02
	#axisError := #InputData.ZSW1_Bit03_Fault;
	#sbFault := #InputData.ZSW1_Bit03_Fault; // 同Bit03
	#axisWarn := #InputData.ZSW1_Bit07_Alarm;
	#sbAlarm := #InputData.ZSW1_Bit07_Alarm; // 同Bit07
	#axisPosOk := #InputData.ZSW1_Bit10_TargetReached;
	#axisRef := #InputData.ZSW1_Bit11_HomeSet;
	#axisSpFixed := #InputData.ZSW1_Bit13_SetpointFixed;
	#sbAccel := #InputData.ZSW1_Bit14_AxisAccel;
	#sbDecel := #InputData.ZSW1_Bit15_AxisDecel;
	#sbBusy := #InputData.ZSW1_Bit02_Enabled; // 使用Enabled作为Busy指示

	// 运动方向
	// #sbFWD := #InputData.POS_ZSW2_Bit04_Forward;
	// #sbBWD := #InputData.POS_ZSW2_Bit05_Backward;

	// 实际值
	#actVelocity := #InputData.VIST;
	#actPosition := #InputData.XIST;
	#actMode := #modePos;

	// 警告和故障代码
	#actWarn := #InputData.AlarmCode;
	#actFault := #InputData.FaultCode;
	#lockOut := #InputData.ZSW1_Bit06_Inhibit;

	// 输出赋值
	#status := #swStatus;
END_FUNCTION_BLOCK

FUNCTION "FC_Delay_On_Variant" : Void
{ S7_Optimized_Access := 'TRUE' }
VERSION : 0.1
   VAR_INPUT
      i_CMD_Start : Bool;
      i_CFG_Target : Variant;
      i_Cycle_Count : Int;
   END_VAR

   VAR_OUTPUT
      o_Delay_Finish : Bool;
   END_VAR

   VAR_IN_OUT
      io_Setpoint : Variant;
   END_VAR

   VAR_TEMP
      t_Int : Struct
         Target : Int;
         Setpoint : Int;
      END_STRUCT;
      t_DInt : Struct
         Target : DInt;
         Setpoint : DInt;
      END_STRUCT;
      t_Type_Int_Used : Bool;
      t_Type_DInt_Used : Bool;
   END_VAR


BEGIN
	REGION NETWORK: Init Value
	    #o_Delay_Finish := FALSE;
	    #t_Type_Int_Used := FALSE;
	    #t_Type_DInt_Used := FALSE;
	END_REGION

	REGION NETWORK: Check Type
	    IF TypeOf(#i_CFG_Target) <> TypeOf(#io_Setpoint) THEN
	        RETURN;
	    END_IF;

	    IF TypeOf(#i_CFG_Target) = Int THEN
	        VariantGet(SRC := #i_CFG_Target,
	                   DST => #t_Int.Target);
	        VariantGet(SRC := #io_Setpoint,
	                   DST => #t_Int.Setpoint);
	        #t_Type_Int_Used := TRUE;
	    ELSIF TypeOf(#i_CFG_Target) = DInt THEN
	        VariantGet(SRC := #i_CFG_Target,
	                   DST => #t_DInt.Target);
	        VariantGet(SRC := #io_Setpoint,
	                   DST => #t_DInt.Setpoint);
	        #t_Type_DInt_Used := TRUE;
	    ELSE
	        RETURN;
	    END_IF;
	END_REGION

	REGION NETWORK: Init Timer
	    IF NOT #i_CMD_Start THEN
	        #t_Int.Setpoint := 0;
	        #t_DInt.Setpoint := 0;
	    END_IF;
	END_REGION

	REGION NETWORK: Detect result
	    #o_Delay_Finish := #i_CMD_Start
	    AND ((#t_Type_Int_Used AND #t_Int.Setpoint >= #t_Int.Target)
	    OR (#t_Type_DInt_Used AND #t_DInt.Setpoint >= #t_DInt.Target));
	END_REGION

	REGION NETWORK: Count time value
	    IF #i_CMD_Start THEN
	        IF #t_Type_Int_Used THEN
	            #t_Int.Setpoint := #t_Int.Setpoint + #i_Cycle_Count;
	            IF #t_Int.Setpoint > #t_Int.Target THEN
	                #t_Int.Setpoint := #t_Int.Target;
	            END_IF;
	        ELSIF #t_Type_DInt_Used THEN
	            #t_DInt.Setpoint := #t_DInt.Setpoint + #i_Cycle_Count;
	            IF #t_DInt.Setpoint > #t_DInt.Target THEN
	                #t_DInt.Setpoint := #t_DInt.Target;
	            END_IF;
	        END_IF;
	    END_IF;
	END_REGION

	REGION NETWORK: Write Setpoint
	    IF #t_Type_Int_Used THEN
	        VariantPut(SRC := #t_Int.Setpoint,
	                   DST := #io_Setpoint);
	    ELSIF #t_Type_DInt_Used THEN
	        VariantPut(SRC := #t_DInt.Setpoint,
	                   DST := #io_Setpoint);
	    END_IF;
	END_REGION

END_FUNCTION

FUNCTION "FC_Delay_On_Accumulator_Variant" : Void
{ S7_Optimized_Access := 'TRUE' }
VERSION : 0.1
   VAR_INPUT
      i_CMD_Start : Bool;
      i_Enable_Dly : Bool;
      i_CFG_Target : Variant;
      i_Cycle_Count : Int;
   END_VAR

   VAR_OUTPUT
      o_Delay_Finish : Bool;
   END_VAR

   VAR_IN_OUT
      io_Setpoint : Variant;
   END_VAR

   VAR_TEMP
      t_Int : Struct
         Target : Int;
         Setpoint : Int;
      END_STRUCT;
      t_DInt : Struct
         Target : DInt;
         Setpoint : DInt;
      END_STRUCT;
      t_Type_Int_Used : Bool;
      t_Type_DInt_Used : Bool;
   END_VAR


BEGIN
	REGION NETWORK: Init Value
	    #o_Delay_Finish := FALSE;
	    #t_Type_Int_Used := FALSE;
	    #t_Type_DInt_Used := FALSE;
	END_REGION

	REGION NETWORK: Check Type
	    IF TypeOf(#i_CFG_Target) <> TypeOf(#io_Setpoint) THEN
	        RETURN;
	    END_IF;

	    IF TypeOf(#i_CFG_Target) = Int THEN
	        VariantGet(SRC := #i_CFG_Target,
	                   DST => #t_Int.Target);
	        VariantGet(SRC := #io_Setpoint,
	                   DST => #t_Int.Setpoint);
	        #t_Type_Int_Used := TRUE;
	    ELSIF TypeOf(#i_CFG_Target) = DInt THEN
	        VariantGet(SRC := #i_CFG_Target,
	                   DST => #t_DInt.Target);
	        VariantGet(SRC := #io_Setpoint,
	                   DST => #t_DInt.Setpoint);
	        #t_Type_DInt_Used := TRUE;
	    ELSE
	        RETURN;
	    END_IF;
	END_REGION

	REGION NETWORK: Init Timer
	    IF NOT #i_CMD_Start THEN
	        #t_Int.Setpoint := 0;
	        #t_DInt.Setpoint := 0;
	    END_IF;
	END_REGION

	REGION NETWORK: Detect result
	    #o_Delay_Finish := #i_CMD_Start
	    AND ((#t_Type_Int_Used AND #t_Int.Setpoint >= #t_Int.Target)
	    OR (#t_Type_DInt_Used AND #t_DInt.Setpoint >= #t_DInt.Target));
	END_REGION

	REGION NETWORK: Count time value
	    IF #i_CMD_Start THEN
	        IF #t_Type_Int_Used THEN
	            IF #i_Enable_Dly THEN
	                #t_Int.Setpoint := #t_Int.Setpoint + #i_Cycle_Count;
	            END_IF;
	            IF #t_Int.Setpoint > #t_Int.Target THEN
	                #t_Int.Setpoint := #t_Int.Target;
	            END_IF;
	        ELSIF #t_Type_DInt_Used THEN
	            IF #i_Enable_Dly THEN
	                #t_DInt.Setpoint := #t_DInt.Setpoint + #i_Cycle_Count;
	            END_IF;
	            IF #t_DInt.Setpoint > #t_DInt.Target THEN
	                #t_DInt.Setpoint := #t_DInt.Target;
	            END_IF;
	        END_IF;
	    END_IF;
	END_REGION

	REGION NETWORK: Write Setpoint
	    IF #t_Type_Int_Used THEN
	        VariantPut(SRC := #t_Int.Setpoint,
	                   DST := #io_Setpoint);
	    ELSIF #t_Type_DInt_Used THEN
	        VariantPut(SRC := #t_DInt.Setpoint,
	                   DST := #io_Setpoint);
	    END_IF;
	END_REGION
END_FUNCTION

TYPE "UDT_Global"
TITLE = UDT_Global
VERSION : 0.1
//General runtime variable
//# Block Info
//- Title:            UDT_Global
//- Comment/Function: General runtime variable
//- Library/Family:   APS
//- Author:           Jay Liu
//- Tested with:      ---
//- Engineering:      TIA Portal V20
//- Restrictions:     ---
//- Requirements:     ---
//
//# History
// |Version  | Date       | Author                 | Description                   |
// |---------|------------|------------------------|------------------------------ |
// |01.00.00 | 2026-01-22 | Jay Liu                | First released version        |
   STRUCT
      AlwaysOff : Bool;   // FALSE
      AlwaysOn : Bool;   // TRUE
      PLC_Is_Simulated : Bool;   // Indicates that simulated PLC is used
      PLC_1200 : Bool;   // PLC is 1200 series
      PLC_1500 : Bool;   // PLC is 1500 series
      PLC_NoFailsafe : Bool;   // PLC donot support failsafe
      OS_First_Scan : Bool;   // TRUE during 1st. scan after Restart
      OS_New_Year : Bool;   // One-Shot each year
      OS_New_Month : Bool;   // One-Shot each month
      OS_New_Week : Bool;   // One-Shot each week
      OS_New_Day : Bool;   // One-Shot each day
      OS_New_Hour : Bool;   // One-Shot each hour
      OS_New_Minute : Bool;   // One-Shot each minute
      OS_New_Second : Bool;   // One-Shot each second
      Clock_10Hz : Bool;   // 0.05s on, 0.05s off
      Clock_5Hz : Bool;   // 0.01s on, 0.01s off
      Clock_2_5Hz : Bool;   // 0.125s on, 0.125s off
      Clock_2Hz : Bool;   // 0.25s on, 0.25s off
      Clock_1_25Hz : Bool;   // 0.4s on, 0.4s off
      Clock_1Hz : Bool;   // 0.5s on, 0.5s off
      Clock_0_625Hz : Bool;   // 0.8s on, 0.8s off
      Clock_0_5Hz : Bool;   // 1s on, 1s off
      OneShot_0_05sec : Bool;   // One-Shot each 0.05 sec
      OneShot_0_1sec : Bool;   // One-Shot each 0.1 sec
      OneShot_0_2sec : Bool;   // One-Shot each 0.2sec
      OneShot_0_25sec : Bool;   // One-Shot each 0.25 sec
      OneShot_0_5sec : Bool;   // One-Shot each 0.5 sec
      OneShot_0_8sec : Bool;   // One-Shot each 0.8 sec
      OneShot_1sec : Bool;   // One-Shot each 1 sec
      OneShot_2sec : Bool;   // One-Shot each 2 sec
      OB_Prev_Cycle_Time : Int;   // [ms] Passed time in previous PLC cycle
      OB_Average_Cycle_Time : Int;   // [ms] Average passed time in previous PLC cycle
      OB_Min_Cycle_Time : Int := 9999;   // [ms] The minimum passed time in previous PLC cycle
      OB_Max_Cycle_Time : Int;   // [ms] The maximum passed time in previous PLC cycle
      Common_Setting : "UDT_Commen_Setting";
   END_STRUCT;

END_TYPE

DATA_BLOCK "DB_Setting"
TITLE = %version: 544e4e8 % CN: 20
{ S7_Optimized_Access := 'FALSE' }
FAMILY : General
VERSION : 0.0
//History:
//repo_name:     ALLCTTT/VI_TTT
//status:        release-3.7.0.0
//
//All commits of this file:
//
//IssueID            Description                                            By                             CommitDate CommitID
//----------------------------------------------------------------------------------------------------------------------------
//ALLCTTT-272        removed keywords                                       Pascal van Kempen              2020-12-10 544e4e8
//ALLCTTT-272        Revert ALLCTTT-272 - corrected checkin sequence for de Pascal van Kempen              2020-12-10 9d531fb
//ALLCTTT-272        corrected checkin sequence for determining version inf Pascal van Kempen              2020-12-10 ae3fa86
//ALLCTTT-272        Revert ALLCTTT-272 - keywords updates                  Pascal van Kempen              2020-12-10 5a1edb7
//ALLCTTT-272        keywords updates                                       Pascal van Kempen              2020-12-10 8d62c21
//ALLCTTT-272        initial import                                         Pascal van Kempen              2020-12-10 31a6487
//
//This version
//              %date_created: 2020-12-10 17:18:38 +0100 %
//              %release: %
//
//Modification History:                                 By:      Date:     Rev:
//----------------------------------------------------  -------  --------  -----
//ra#31964: Based on 2.15.0.0 version 1.01              nlhhop   14-01-19   2.01
   STRUCT
      Common : "UDT_Commen_Setting";
      SSM : "UDT_SSM_Setting";
      AWCS : "UDT_AWCS_Setting";
      PLC_Log : "UDT_PLC_Log_Setting";
      GC03_CT01 : "UDT_Datalogic_AV900_Setting";
      GC04_CT01 : "UDT_Datalogic_AV900_Setting";
      Tipper01 : "UDT_Tipper_Setting";
      ECH01 : "UDT_Echelon_Setting";
      RLS01 : "UDT_RLS_Setting";
      Tipper02 : "UDT_Tipper_Setting";
      ECH02 : "UDT_Echelon_Setting";
      RLS02 : "UDT_RLS_Setting";
      SG : "UDT_Merge_Singulator_Setting";
      IBST : "UDT_NBS_Setting";
      ADTA : "UDT_ADTA_Setting";
      GC01_A01 : "UDT_IOLink_Master_Setting";
      GC01_A02 : "UDT_IOLink_Master_Setting";
      GC01_A03 : "UDT_IOLink_Master_Setting";
      GC01_A04 : "UDT_IOLink_Master_Setting";
      GC01_A05 : "UDT_IOLink_Master_Setting";
      GC02_A01 : "UDT_IOLink_Master_Setting";
      GC02_A02 : "UDT_IOLink_Master_Setting";
      GC02_A03 : "UDT_IOLink_Master_Setting";
      GC03_A01 : "UDT_IOLink_Master_Setting";
      GC03_A02 : "UDT_IOLink_Master_Setting";
      GC03_A03 : "UDT_IOLink_Master_Setting";
      GC03_A04 : "UDT_IOLink_Master_Setting";
      GC03_A05 : "UDT_IOLink_Master_Setting";
      GC03_A06 : "UDT_IOLink_Master_Setting";
      GC04_A01 : "UDT_IOLink_Master_Setting";
      GC04_A02 : "UDT_IOLink_Master_Setting";
      GC04_A03 : "UDT_IOLink_Master_Setting";
      GC05_A01 : "UDT_IOLink_Master_Setting";
      GC06_A01 : "UDT_IOLink_Master_Setting";
      GC07_A01 : "UDT_IOLink_Master_Setting";
      GC01_FB01 : "UDT_Conv_G115D_Setting";
      GC01_FB02 : "UDT_Conv_G115D_Setting";
      GC01_FB03 : "UDT_Conv_G115D_Setting";
      GC01_FB03_Track : "UDT_Track_Setting";
      GC01_FB04 : "UDT_Conv_S210_Setting";
      GC01_FB04_Track : "UDT_Track_Setting";
      GC01_FB05 : "UDT_Conv_S210_Setting";
      GC01_FB05_Track : "UDT_Track_Setting";
      DT01 : "UDT_Conv_SWS_Setting";
      GC01_RC06_Track : "UDT_Track_Setting";
      GC01_RC06 : "UDT_Conv_MultiControl_Setting";
      GC01_FB07 : "UDT_Conv_G115D_Setting";
      GC01_FB08 : "UDT_Conv_G115D_Setting";
      GC01_RC09_Track : "UDT_Track_Setting";
      GC01_RC09 : "UDT_Conv_MultiControl_Setting";
      GC01_RC10 : "UDT_Conv_MultiControl_Setting";
      GC01_RC40 : "UDT_Conv_MultiControl_Setting";
      GC01_SK11 : "UDT_Conv_G115D_Setting";
      GC01_FB12 : "UDT_Conv_S210_Setting";
      GC01_FB13 : "UDT_Conv_S210_Setting";
      GC01_FB14 : "UDT_Conv_S210_Setting";
      GC01_FB15 : "UDT_Conv_G115D_Setting";
      GC01_FB16 : "UDT_Conv_G115D_Setting";
      GC01_FB17 : "UDT_Conv_G115D_Setting";
      GC01_FB18 : "UDT_Conv_G115D_Setting";
      GC01_FB19 : "UDT_Conv_G115D_Setting";
      GC01_FB20 : "UDT_Conv_G115D_Setting";
      GC01_FB21 : "UDT_Conv_G115D_Setting";
      GC01_FB22 : "UDT_Conv_G115D_Setting";
      GC01_FB23 : "UDT_Conv_G115D_Setting";
      GC01_FB24 : "UDT_Conv_G115D_Setting";
      GC01_FB25 : "UDT_Conv_G115D_Setting";
      GC01_FB26 : "UDT_Conv_G115D_Setting";
      GC01_FB27 : "UDT_Conv_G115D_Setting";
      GC01_FB28 : "UDT_Conv_S210_Setting";
      GC01_FB29 : "UDT_Conv_S210_Setting";
      GC01_FB30 : "UDT_Conv_S210_Setting";
      GC01_FB31 : "UDT_Conv_S210_Setting";
      GC01_FB32 : "UDT_Conv_G115D_Setting";
      GC02_FB01 : "UDT_Conv_G115D_Setting";
      GC02_FB02 : "UDT_Conv_G115D_Setting";
      GC02_FB03 : "UDT_Conv_S210_Setting";
      GC02_FB03_Track : "UDT_Track_Setting";
      GC02_FB04 : "UDT_Conv_S210_Setting";
      GC02_FB04_Track : "UDT_Track_Setting";
      DT02 : "UDT_Conv_SWS_Setting";
      GC02_RC05_Track : "UDT_Track_Setting";
      GC02_RC05 : "UDT_Conv_MultiControl_Setting";
      GC02_FB06 : "UDT_Conv_G115D_Setting";
      GC02_FB07 : "UDT_Conv_G115D_Setting";
      GC02_FB08_Track : "UDT_Track_Setting";
      GC02_FB08 : "UDT_Conv_G115D_Setting";
      GC02_FB09 : "UDT_Conv_G115D_Setting";
      GC02_FB10 : "UDT_Conv_G115D_Setting";
      GC02_FB11 : "UDT_Conv_G115D_Setting";
      GC02_FB12 : "UDT_Conv_G115D_Setting";
      GC02_FB13 : "UDT_Conv_G115D_Setting";
      GC02_FB14 : "UDT_Conv_G115D_Setting";
      GC02_SK15 : "UDT_Conv_G115D_Setting";
      GC02_FB16 : "UDT_Conv_S210_Setting";
      GC02_FB17 : "UDT_Conv_S210_Setting";
      GC02_FB18 : "UDT_Conv_S210_Setting";
      GC03_RC01 : "UDT_Conv_MultiControl_Setting";
      GC03_RC40 : "UDT_Conv_MultiControl_Setting";
      GC03_RC02 : "UDT_Conv_MultiControl_Setting";
      GC03_RC03 : "UDT_Conv_MultiControl_Setting";
      GC03_RC41 : "UDT_Conv_MultiControl_Setting";
      GC03_RC04 : "UDT_Conv_MultiControl_Setting";
      GC03_HB05_Merge : "UDT_Merge_2_To_1_Setting";
      GC03_HB05 : "UDT_Conv_Multiple_S210_Setting";
      GC03_FB06 : "UDT_Conv_G115D_Setting";
      GC03_FB42 : "UDT_Conv_G115D_Setting";
      GC03_FB07 : "UDT_Conv_G115D_Setting";
      GC03_FB08_Track : "UDT_Track_Setting";
      GC03_FB08 : "UDT_Conv_G115D_Setting";
      GC03_FB09_Track : "UDT_Track_Setting";
      GC03_FB09 : "UDT_Conv_G115D_Setting";
      GC03_FB10 : "UDT_Conv_S210_Setting";
      GC03_FB11_Track : "UDT_Track_Setting";
      GC03_FB11 : "UDT_Conv_S210_Setting";
      DT03 : "UDT_Conv_SWS_Setting";
      GC03_RC12_Track : "UDT_Track_Setting";
      GC03_RC12 : "UDT_Conv_MultiControl_Setting";
      GC03_FB13 : "UDT_Conv_G115D_Setting";
      GC03_FB14 : "UDT_Conv_S210_Setting";
      GC03_FB15 : "UDT_Conv_S210_Setting";
      GC03_FB16 : "UDT_Conv_S210_Setting";
      GC03_FB17 : "UDT_Conv_S210_Setting";
      GC03_FB18 : "UDT_Conv_G115D_Setting";
      GC03_RC19 : "UDT_Conv_G115D_Setting";
      GC03_RC20 : "UDT_Conv_MultiControl_Setting";
      GC03_FB21_Accmulation : "UDT_Accmulation_Setting";
      GC03_FB21 : "UDT_Conv_G115D_Setting";
      GC03_FB22 : "UDT_Conv_G115D_Setting";
      GC03_FB23 : "UDT_Conv_G115D_Setting";
      GC03_FB24 : "UDT_Conv_G115D_Setting";
      GC03_FB25 : "UDT_Conv_G115D_Setting";
      GC03_FB26 : "UDT_Conv_G115D_Setting";
      GC03_FB27 : "UDT_Conv_G115D_Setting";
      GC03_FB28 : "UDT_Conv_G115D_Setting";
      GC03_FB29 : "UDT_Conv_G115D_Setting";
      GC03_FB30 : "UDT_Conv_G115D_Setting";
      GC03_FB31 : "UDT_Conv_G115D_Setting";
      GC03_FB32_Infeed : "UDT_Induct_On_Gap_Setting";
      GC03_FB32 : "UDT_Conv_G115D_Setting";
      GC03_RC33_Track : "UDT_Track_Setting";
      GC03_RC33 : "UDT_Conv_Dual_G115D_Setting";
      GC04_FB04 : "UDT_Conv_G115D_Setting";
      GC04_FB05 : "UDT_Conv_G115D_Setting";
      GC04_FB06 : "UDT_Conv_G115D_Setting";
      GC04_FB07 : "UDT_Conv_G115D_Setting";
      GC04_FB08 : "UDT_Conv_G115D_Setting";
      GC04_FB09_Track : "UDT_Track_Setting";
      GC04_FB09 : "UDT_Conv_G115D_Setting";
      GC04_FB10 : "UDT_Conv_S210_Setting";
      GC04_FB11_Track : "UDT_Track_Setting";
      GC04_FB11 : "UDT_Conv_S210_Setting";
      DT04 : "UDT_Conv_SWS_Setting";
      GC04_CH01 { S7_SetPoint := 'False'} : "UDT_Chute_Setting";
      GC04_FB12 : "UDT_Conv_G115D_Setting";
      GC04_FB13_Track : "UDT_Track_Setting";
      GC04_FB13 : "UDT_Conv_G115D_Setting";
      GC04_FB14 : "UDT_Conv_G115D_Setting";
      GC04_FB15 : "UDT_Conv_G115D_Setting";
      GC04_FB16 : "UDT_Conv_G115D_Setting";
      GC04_FB17 : "UDT_Conv_G115D_Setting";
      GC04_FB18 : "UDT_Conv_G115D_Setting";
      GC04_FB19 : "UDT_Conv_G115D_Setting";
      GC04_RC20 : "UDT_Conv_MultiControl_Setting";
      GC04_RC21_Track : "UDT_Track_Setting";
      GC04_RC21 : "UDT_Conv_Dual_G115D_Setting";
      GC05_RC01 : "UDT_Conv_MultiControl_Setting";
      GC05_RC02 : "UDT_Conv_MultiControl_Setting";
      GC05_RC03 : "UDT_Conv_MultiControl_Setting";
      GC05_RC10 : "UDT_Conv_MultiControl_Setting";
      GC05_FB04 : "UDT_Conv_G115D_Setting";
      GC05_FB05 : "UDT_Conv_G115D_Setting";
      GC05_RC06 : "UDT_Conv_MultiControl_Setting";
      GC05_RC07 : "UDT_Conv_G115D_Setting";
      GC06_RC01 : "UDT_Conv_MultiControl_Setting";
      GC06_FB02 : "UDT_Conv_G115D_Setting";
      GC06_FB03 : "UDT_Conv_G115D_Setting";
      GC06_RC04_Merge : "UDT_Merge_3_To_1_Setting";
      GC06_RC04 : "UDT_Conv_Triple_G115D_Setting";
      GC06_FB05 : "UDT_Conv_G115D_Setting";
      GC06_FB06 : "UDT_Conv_G115D_Setting";
      GC06_FB07 : "UDT_Conv_G115D_Setting";
      GC06_SK08 : "UDT_Conv_G115D_Setting";
      GC07_CH01 { S7_SetPoint := 'False'} : "UDT_Chute_Setting";
      GC07_FB01 : "UDT_Conv_G115D_Setting";
      GC07_RC02 : "UDT_Conv_Dual_G115D_Setting";
      GC07_RC03 : "UDT_Conv_MultiControl_Setting";
      GC07_RC04 : "UDT_Conv_MultiControl_Setting";
      GC07_RC05 : "UDT_Conv_MultiControl_Setting";
      GC07_RC06 : "UDT_Conv_MultiControl_Setting";
      GC07_RC10 : "UDT_Conv_MultiControl_Setting";
      GC07_RC07 : "UDT_Conv_MultiControl_Setting";
      GC07_RC08 : "UDT_Conv_MultiControl_Setting";
      GC07_RC11 : "UDT_Conv_MultiControl_Setting";
      GC07_CH02 { S7_SetPoint := 'False'} : "UDT_Chute_Setting";
      GC07_FB09 : "UDT_Conv_G115D_Setting";
   END_STRUCT;


BEGIN
   Common.Disable_Energy_Saving := TRUE;
   SSM.StartUp_Indication_Time := 5;
   SSM.Restart_Indication_Time := 5;
   SSM.ControlStop_Time := 60;
   AWCS.InterfaceId := 64;
   AWCS.ID_Range := 1;
   AWCS.LocalPort := 5001;
   PLC_Log.Connection.ID := 10;
   GC03_CT01.Scanner_ID := 'GC03_CT01';
   GC04_CT01.Scanner_ID := 'GC04_CT01';
   ECH01.StartUp_Delay := 2000;
   SG.StartUp_Delay := 1000;
   IBST.StartUp_Delay := 3000;
   DT01.Decision.Straight_Destination := 3;
   DT01.Decision.Left_Destination := 1;
   DT01.Decision.Right_Destination := 2;
   DT01.Decision.High_Priority := 2;
   DT01.Decision.Middle_Priority := 4;
   DT01.Decision.Low_Priority := 8;
   DT01.Decision.Default_Direction := 8;
   DT01.Decision.Destination_Invalid.Enable := TRUE;
   DT01.Decision.Destination_Invalid.Preferred_Direction := 16#0008;
   DT01.Decision.No_Destination.Enable := TRUE;
   DT01.Decision.No_Destination.Preferred_Direction := 16#0008;
   DT01.Decision.Gap_Error.Preferred_Direction := 16#0008;
   DT01.Decision.Diemension_Error.Enable := TRUE;
   DT01.Decision.Diemension_Error.Threshold := 120;
   DT01.Decision.Diemension_Error.Preferred_Direction := 16#0008;
   DT01.Decision.Dir_Fault_Straight.Enable := TRUE;
   DT01.Decision.Dir_Fault_Straight.Disallowed_Direction := 16#0002;
   DT01.Decision.Dir_Fault_Left.Enable := TRUE;
   DT01.Decision.Dir_Fault_Left.Disallowed_Direction := 16#0004;
   DT01.Decision.Dir_Fault_Right.Disallowed_Direction := 16#0008;
   DT01.Decision.Dir_Disabled_Straight.Enable := TRUE;
   DT01.Decision.Dir_Disabled_Straight.Disallowed_Direction := 16#0002;
   DT01.Decision.Dir_Disabled_Left.Enable := TRUE;
   DT01.Decision.Dir_Disabled_Left.Disallowed_Direction := 16#0004;
   DT01.Decision.Dir_Disabled_Right.Disallowed_Direction := 16#0008;
   DT01.Decision.Dir_Full_Straight.Enable := TRUE;
   DT01.Decision.Dir_Full_Straight.Disallowed_Direction := 16#0002;
   DT01.Decision.Dir_Full_Left.Enable := TRUE;
   DT01.Decision.Dir_Full_Left.Disallowed_Direction := 16#0004;
   DT01.Decision.Dir_Full_Right.Disallowed_Direction := 16#0008;
   DT01.Decision.No_Read.Enable := TRUE;
   DT01.Decision.No_Read.Preferred_Direction := 16#0008;
   DT01.Decision.No_Code.Enable := TRUE;
   DT01.Decision.No_Code.Preferred_Direction := 16#0008;
   DT01.Decision.Multi_Read.Enable := TRUE;
   DT01.Decision.Multi_Read.Preferred_Direction := 16#0008;
   DT01.Decision.Unexpected_Item.Enable := TRUE;
   DT01.Decision.Unexpected_Item.Preferred_Direction := 16#0008;
   DT01.Divert.Fixed_Ratio_Left := 1;
   DT01.Divert.Fixed_Ratio_Right := 1;
   DT01.Divert.First_Group_Action_Delay := 35;
   DT01.Divert.Group2_Action_Delay := 16;
   DT01.Divert.Group3_Action_Delay := 16;
   DT01.Divert.Group4_Action_Delay := 16;
   DT01.Divert.Group5_Action_Delay := 17;
   DT01.Divert.Group6_Action_Delay := 17;
   DT01.Divert.Group7_Action_Delay := 17;
   DT01.Divert.Group8_Action_Delay := 17;
   DT01.Divert.Group9_Action_Delay := 17;
   DT01.Base_Conveyor.Delay_Dieback := 0;
   DT01.Base_Conveyor.Delay_Startup := 0;
   DT01.Base_Conveyor.Delay_Cascade_Startup := 0;
   DT01.Base_Conveyor.Slave_Mode := TRUE;
   DT01.Hardware.Servo_U401.Left_Position_Setpoint := -25;
   DT01.Hardware.Servo_U411.Left_Position_Setpoint := -40;
   DT01.Hardware.Servo_U421.Left_Position_Setpoint := -55;
   DT01.Hardware.Servo_U431.Left_Position_Setpoint := -55;
   DT01.Hardware.Servo_U441.Left_Position_Setpoint := -55;
   DT01.Hardware.Servo_U451.Left_Position_Setpoint := -55;
   DT01.Hardware.Servo_U461.Left_Position_Setpoint := -55;
   DT01.Hardware.Servo_U471.Left_Position_Setpoint := -55;
   DT01.Hardware.Servo_U481.Left_Position_Setpoint := -55;
   GC01_RC06.Hardware_U01.Speed1 := 1200;
   GC01_RC06.Hardware_U01.RefSpeed := 1390;
   GC01_RC06.Hardware_U01.RD1_Motor_Number := 1;
   GC01_RC06.Hardware_U01.RD2_Motor_Number := 2;
   GC01_FB08.Base_Conveyor.Slave_Mode := TRUE;
   GC01_RC09_Track.Measure_Length := TRUE;
   GC01_RC09_Track.Localtion := 'GC01_RC09';
   GC01_RC09.Base_Conveyor.Slave_Mode := TRUE;
   GC01_RC09.Hardware_U01.Speed1 := 1200;
   GC01_RC09.Hardware_U01.RefSpeed := 1390;
   GC01_RC09.Hardware_U01.RD1_Motor_Number := 1;
   GC01_RC09.Hardware_U01.RD2_Motor_Number := 2;
   GC01_RC10.Base_Conveyor.Slave_Mode := TRUE;
   GC01_RC10.Hardware_U01.Speed1 := 1000;
   GC01_RC10.Hardware_U01.RefSpeed := 1390;
   GC01_RC10.Hardware_U01.RD1_Motor_Number := 1;
   GC01_RC10.Hardware_U01.RD2_Motor_Number := 2;
   GC01_RC10.Hardware_U01.RD3_Motor_Number := 3;
   GC01_RC40.Hardware_U01.Speed1 := 1000;
   GC01_RC40.Hardware_U01.RefSpeed := 1390;
   GC01_RC40.Hardware_U01.RD4_Motor_Number := 1;
   GC01_FB15.Hardware.Speed1 := 2000;
   GC01_FB16.Hardware.Speed1 := 2000;
   GC01_FB17.Hardware.Speed1 := 2000;
   GC01_FB18.Hardware.Speed1 := 2000;
   GC01_FB19.Hardware.Speed1 := 2000;
   GC01_FB20.Hardware.Speed1 := 2000;
   GC01_FB21.Hardware.Speed1 := 2000;
   GC01_FB22.Hardware.Speed1 := 2000;
   GC01_FB23.Hardware.Speed1 := 2000;
   GC01_FB24.Hardware.Speed1 := 2000;
   GC01_FB25.Hardware.Speed1 := 2000;
   GC01_FB26.Hardware.Speed1 := 2000;
   GC01_FB27.Hardware.Speed1 := 2000;
   GC01_FB28.Hardware.Speed1 := 2000;
   GC01_FB29.Hardware.Speed1 := 2000;
   GC01_FB30.Hardware.Speed1 := 2000;
   GC01_FB31.Hardware.Speed1 := 2000;
   GC01_FB32.Hardware.Speed1 := 2000;
   GC02_RC05.Hardware_U01.Speed1 := 1200;
   GC02_RC05.Hardware_U01.RefSpeed := 1390;
   GC02_RC05.Hardware_U01.RD1_Motor_Number := 1;
   GC02_RC05.Hardware_U01.RD2_Motor_Number := 2;
   GC03_RC01.Base_Conveyor.Slave_Mode := TRUE;
   GC03_RC01.Hardware_U01.Speed1 := 500;
   GC03_RC01.Hardware_U01.RefSpeed := 1000;
   GC03_RC01.Hardware_U01.RD1_Motor_Number := 1;
   GC03_RC01.Hardware_U01.RD2_Motor_Number := 2;
   GC03_RC40.Base_Conveyor.Slave_Mode := TRUE;
   GC03_RC40.Hardware_U01.Speed1 := 500;
   GC03_RC40.Hardware_U01.RefSpeed := 1000;
   GC03_RC40.Hardware_U01.RD3_Motor_Number := 1;
   GC03_RC40.Hardware_U01.RD4_Motor_Number := 2;
   GC03_RC02.PE1.Handover_Offset := 200;
   GC03_RC02.Hardware_U01.Speed1 := 500;
   GC03_RC02.Hardware_U01.RefSpeed := 1000;
   GC03_RC02.Hardware_U01.RD1_Motor_Number := 1;
   GC03_RC02.Hardware_U01.RD2_Motor_Number := 2;
   GC03_RC02.Hardware_U01.RD3_Motor_Number := 3;
   GC03_RC03.Base_Conveyor.Slave_Mode := TRUE;
   GC03_RC03.Hardware_U01.Speed1 := 500;
   GC03_RC03.Hardware_U01.RefSpeed := 1000;
   GC03_RC03.Hardware_U01.RD1_Motor_Number := 1;
   GC03_RC03.Hardware_U01.RD2_Motor_Number := 2;
   GC03_RC41.Base_Conveyor.Slave_Mode := TRUE;
   GC03_RC41.Hardware_U01.Speed1 := 500;
   GC03_RC41.Hardware_U01.RefSpeed := 1000;
   GC03_RC41.Hardware_U01.RD3_Motor_Number := 1;
   GC03_RC41.Hardware_U01.RD4_Motor_Number := 2;
   GC03_RC04.PE1.Handover_Offset := 200;
   GC03_RC04.Hardware_U01.Speed1 := 500;
   GC03_RC04.Hardware_U01.RefSpeed := 1000;
   GC03_RC04.Hardware_U01.RD1_Motor_Number := 1;
   GC03_RC04.Hardware_U01.RD2_Motor_Number := 2;
   GC03_RC04.Hardware_U01.RD3_Motor_Number := 3;
   GC03_HB05_Merge.Line1_Infeed_Delay := 500;
   GC03_HB05_Merge.Line2_Infeed_Delay := 500;
   GC03_FB06.Base_Conveyor.Slave_Mode := TRUE;
   GC03_FB07.Base_Conveyor.Slave_Mode := TRUE;
   GC03_FB08_Track.Measure_Length := TRUE;
   GC03_FB08_Track.Package_Range := 3;
   GC03_FB08_Track.Localtion := 'GC03_FB08';
   GC03_FB08.Base_Conveyor.Slave_Mode := TRUE;
   GC03_FB09_Track.Measure_Length := TRUE;
   GC03_FB09_Track.Update_Position := 5450;
   GC03_FB09_Track.Package_Range := 3;
   GC03_FB09_Track.Localtion := 'GC03_FB09';
   GC03_FB09.Base_Conveyor.Slave_Mode := TRUE;
   GC03_FB10.Base_Conveyor.Slave_Mode := TRUE;
   GC03_FB11_Track.Update_Position := 7900;
   GC03_FB11_Track.Package_Range := 3;
   GC03_FB11_Track.Localtion := 'GC03_FB11';
   GC03_FB11.Base_Conveyor.Slave_Mode := TRUE;
   DT03.Decision.Decision_Position := 8100;
   DT03.Decision.Straight_Destination := 7;
   DT03.Decision.Left_Destination := 8;
   DT03.Decision.Right_Destination := 9;
   DT03.Decision.Destination_Invalid.Enable := TRUE;
   DT03.Decision.Destination_Invalid.Preferred_Direction := 16#08;
   DT03.Decision.No_Destination.Enable := TRUE;
   DT03.Decision.No_Destination.Preferred_Direction := 16#08;
   DT03.Decision.Diemension_Error.Enable := TRUE;
   DT03.Decision.Diemension_Error.Threshold := 1200;
   DT03.Decision.Diemension_Error.Preferred_Direction := 16#08;
   DT03.Decision.Throughput_Limit_Straight.Enable := TRUE;
   DT03.Decision.Throughput_Limit_Straight.Preferred_Direction := 16#08;
   DT03.Decision.Throughput_Limit_Left.Enable := TRUE;
   DT03.Decision.Throughput_Limit_Left.Preferred_Direction := 16#08;
   DT03.Decision.Dir_Fault_Straight.Enable := TRUE;
   DT03.Decision.Dir_Fault_Straight.Preferred_Direction := 16#08;
   DT03.Decision.Dir_Fault_Left.Enable := TRUE;
   DT03.Decision.Dir_Fault_Left.Preferred_Direction := 16#08;
   DT03.Decision.Dir_Disabled_Straight.Enable := TRUE;
   DT03.Decision.Dir_Disabled_Straight.Preferred_Direction := 16#08;
   DT03.Decision.Dir_Disabled_Left.Enable := TRUE;
   DT03.Decision.Dir_Disabled_Left.Preferred_Direction := 16#08;
   DT03.Decision.Dir_Full_Straight.Enable := TRUE;
   DT03.Decision.Dir_Full_Straight.Preferred_Direction := 16#08;
   DT03.Decision.Dir_Full_Left.Enable := TRUE;
   DT03.Decision.Dir_Full_Left.Preferred_Direction := 16#08;
   DT03.Base_Conveyor.Slave_Mode := TRUE;
   GC03_RC12_Track.Update_Position := 11040;
   GC03_RC12_Track.Package_Range := 3;
   GC03_RC12_Track.Localtion := 'GC03_RC12';
   GC03_RC12.Hardware_U01.Speed1 := 1200;
   GC03_RC12.Hardware_U01.RefSpeed := 1390;
   GC03_RC12.Hardware_U01.RD2_Motor_Number := 1;
   GC03_RC12.Hardware_U01.RD3_Motor_Number := 2;
   GC03_FB13.PE1.Shifting_Offset := 1300;
   GC03_FB14.PE1.Shifting_Offset := 900;
   GC03_FB14.PE1.Handover_Offset := 500;
   GC03_FB15.PE1.Shifting_Offset := 900;
   GC03_FB15.PE1.Handover_Offset := 500;
   GC03_FB15.Flow_Control.Minimum_Head_To_Head := 1500;
   GC03_FB16.PE1.Shifting_Offset := 900;
   GC03_FB16.PE1.Handover_Offset := 500;
   GC03_FB16.Flow_Control.Minimum_Head_To_Head := 1500;
   GC03_FB17.PE1.Shifting_Offset := 900;
   GC03_FB17.PE1.Handover_Offset := 500;
   GC03_FB17.Flow_Control.Minimum_Head_To_Head := 1500;
   GC03_FB18.PE1.Shifting_Offset := 1100;
   GC03_FB18.PE1.Handover_Offset := 600;
   GC03_FB18.Flow_Control.Minimum_Head_To_Head := 1500;
   GC03_RC20.Base_Conveyor.Slave_Mode := TRUE;
   GC03_RC20.Hardware_U01.Speed1 := 1390;
   GC03_RC20.Hardware_U01.RefSpeed := 1390;
   GC03_RC20.Hardware_U01.RD1_Motor_Number := 1;
   GC03_RC20.Hardware_U02.Speed1 := 1390;
   GC03_RC20.Hardware_U02.RefSpeed := 1390;
   GC03_RC20.Hardware_U02.RD1_Motor_Number := 2;
   GC03_RC20.Hardware_U02.RD2_Motor_Number := 3;
   GC03_RC20.Hardware_U02.RD3_Motor_Number := 4;
   GC03_RC20.Hardware_U02.RD4_Motor_Number := 5;
   GC03_FB21_Accmulation.Gap := 700;
   GC03_FB21_Accmulation.Cleanup_Distance := 10000;
   GC03_FB21_Accmulation.Waiting_Timeout := 30;
   GC03_FB21_Accmulation.Max_Count := 99;
   GC03_FB21.PE1.Shifting_Offset := 400;
   GC03_FB21.PE1.Handover_Offset := 400;
   GC03_FB21.Base_Conveyor.Delay_Startup := 50;
   GC03_FB22.Base_Conveyor.Slave_Mode := TRUE;
   GC03_FB23.PE1.Shifting_Offset := 1300;
   GC03_FB23.PE1.Handover_Offset := 400;
   GC03_FB24.PE1.Handover_Offset := 300;
   GC03_FB25.PE1.Handover_Offset := 300;
   GC03_FB26.PE1.Handover_Offset := 300;
   GC03_FB27.PE1.Handover_Offset := 300;
   GC03_FB28.PE1.Handover_Offset := 300;
   GC03_FB29.Base_Conveyor.Slave_Mode := TRUE;
   GC03_FB30.PE1.Shifting_Offset := 300;
   GC03_FB30.PE1.Handover_Offset := 200;
   GC03_FB31.PE1.Shifting_Offset := 650;
   GC03_FB31.PE1.Handover_Offset := 400;
   GC03_FB31.Flow_Control.Minimum_Head_To_Head := 1200;
   GC03_FB32_Infeed.Induct_Position := 1850;
   GC03_FB32_Infeed.Gap_Length := 300;
   GC03_FB32_Infeed.Max_Item_Length := 1000;
   GC03_FB32.PE1.Shifting_Offset := 650;
   GC03_FB32.PE1.Handover_Offset := 400;
   GC03_FB32.Flow_Control.Minimum_Head_To_Head := 1200;
   GC03_RC33_Track.Update_Position := 5100;
   GC03_RC33_Track.Localtion := 'GC01_RC33';
   GC04_RC20.Hardware_U01.Speed1 := 1200;
   GC04_RC20.Hardware_U01.RefSpeed := 1390;
   GC04_RC20.Hardware_U01.RD1_Motor_Number := 1;
   GC04_RC20.Hardware_U01.RD2_Motor_Number := 2;
   GC05_RC01.Base_Conveyor.Slave_Mode := TRUE;
   GC05_RC01.Hardware_U01.Speed1 := 1390;
   GC05_RC01.Hardware_U01.RefSpeed := 1390;
   GC05_RC01.Hardware_U01.RD1_Motor_Number := 1;
   GC05_RC01.Hardware_U01.RD2_Motor_Number := 2;
   GC05_RC01.Hardware_U01.RD3_Motor_Number := 3;
   GC05_RC01.Hardware_U01.RD4_Motor_Number := 4;
   GC05_RC01.Hardware_U02.Speed1 := 1390;
   GC05_RC01.Hardware_U02.RefSpeed := 1390;
   GC05_RC01.Hardware_U02.RD4_Motor_Number := 5;
   GC05_RC02.PE1.Shifting_Offset := 1000;
   GC05_RC02.PE1.Handover_Offset := 300;
   GC05_RC02.Hardware_U01.Speed1 := 1200;
   GC05_RC02.Hardware_U01.RefSpeed := 1390;
   GC05_RC02.Hardware_U01.RD1_Motor_Number := 1;
   GC05_RC02.Hardware_U01.RD2_Motor_Number := 2;
   GC05_RC02.Hardware_U01.RD3_Motor_Number := 3;
   GC05_RC02.Hardware_U02.Speed1 := 1200;
   GC05_RC02.Hardware_U02.RefSpeed := 1390;
   GC05_RC02.Hardware_U02.RD1_Motor_Number := 4;
   GC05_RC02.Hardware_U02.RD2_Motor_Number := 5;
   GC05_RC02.Hardware_U02.RD3_Motor_Number := 6;
   GC05_RC02.Hardware_U02.RD4_Motor_Number := 7;
   GC05_RC02.Hardware_U03.Speed1 := 1200;
   GC05_RC02.Hardware_U03.RefSpeed := 1390;
   GC05_RC02.Hardware_U03.RD1_Motor_Number := 8;
   GC05_RC02.Hardware_U03.RD2_Motor_Number := 9;
   GC05_RC02.Hardware_U03.RD3_Motor_Number := 10;
   GC05_RC02.Hardware_U03.RD4_Motor_Number := 11;
   GC05_RC02.Hardware_U04.Speed1 := 1200;
   GC05_RC02.Hardware_U04.RefSpeed := 1390;
   GC05_RC02.Hardware_U04.RD1_Motor_Number := 12;
   GC05_RC03.Flow_Control.Minimum_Head_To_Head := 1500;
   GC05_RC03.Base_Conveyor.Slave_Mode := TRUE;
   GC05_RC03.Hardware_U01.Speed1 := 1200;
   GC05_RC03.Hardware_U01.RefSpeed := 1390;
   GC05_RC03.Hardware_U01.RD2_Motor_Number := 1;
   GC05_RC10.PE1.Shifting_Offset := 600;
   GC05_RC10.PE1.Handover_Offset := 500;
   GC05_RC10.Hardware_U01.Speed1 := 1200;
   GC05_RC10.Hardware_U01.RefSpeed := 1390;
   GC05_RC10.Hardware_U01.RD3_Motor_Number := 1;
   GC05_FB04.PE1.Shifting_Offset := 3500;
   GC05_FB04.PE1.Handover_Offset := 500;
   GC05_FB04.Base_Conveyor.Slave_Mode := TRUE;
   GC05_FB05.Base_Conveyor.Slave_Mode := TRUE;
   GC05_RC06.PE1.Handover_Offset := 500;
   GC05_RC06.Base_Conveyor.Delay_Dieback := 10;
   GC05_RC06.Hardware_U01.Speed1 := 1390;
   GC05_RC06.Hardware_U01.RefSpeed := 1390;
   GC05_RC06.Hardware_U01.RD1_Motor_Number := 1;
   GC06_RC01.Base_Conveyor.Slave_Mode := TRUE;
   GC06_RC01.Hardware_U01.Speed1 := 1390;
   GC06_RC01.Hardware_U01.RefSpeed := 1390;
   GC06_RC01.Hardware_U01.RD1_Motor_Number := 1;
   GC06_RC01.Hardware_U02.Speed1 := 1390;
   GC06_RC01.Hardware_U02.RefSpeed := 1390;
   GC06_RC01.Hardware_U02.RD1_Motor_Number := 2;
   GC06_RC01.Hardware_U02.RD2_Motor_Number := 3;
   GC06_RC01.Hardware_U02.RD3_Motor_Number := 4;
   GC06_RC01.Hardware_U02.RD4_Motor_Number := 5;
   GC06_FB02.PE1.Shifting_Offset := 1200;
   GC06_FB02.PE1.Handover_Offset := 500;
   GC06_FB03.PE1.Shifting_Offset := 1700;
   GC06_FB03.PE1.Handover_Offset := 500;
   GC06_RC04_Merge.Line1_Infeed_Delay := 500;
   GC06_RC04_Merge.Line1_Waiting_Delay := 1500;
   GC06_RC04_Merge.Line2_Infeed_Delay := 500;
   GC06_RC04_Merge.Line2_Waiting_Delay := 1500;
   GC06_RC04_Merge.Line3_Infeed_Delay := 500;
   GC06_RC04_Merge.Line3_Waiting_Delay := 1000;
   GC06_FB06.Hardware.Speed1 := 1000;
   GC06_FB07.Hardware.Speed1 := 800;
   GC06_SK08.Hardware.Speed1 := 600;
   GC07_RC03.Hardware_U01.Speed1 := 500;
   GC07_RC03.Hardware_U01.RefSpeed := 1000;
   GC07_RC03.Hardware_U01.RD1_Motor_Number := 1;
   GC07_RC04.Hardware_U01.Speed1 := 500;
   GC07_RC04.Hardware_U01.RefSpeed := 1000;
   GC07_RC04.Hardware_U01.RD2_Motor_Number := 1;
   GC07_RC04.Hardware_U01.RD3_Motor_Number := 2;
   GC07_RC04.Hardware_U01.RD4_Motor_Number := 3;
   GC07_RC04.Hardware_U02.Speed1 := 500;
   GC07_RC04.Hardware_U02.RefSpeed := 1000;
   GC07_RC04.Hardware_U02.RD1_Motor_Number := 4;
   GC07_RC04.Hardware_U02.RD2_Motor_Number := 5;
   GC07_RC04.Hardware_U02.RD3_Motor_Number := 6;
   GC07_RC04.Hardware_U02.RD4_Motor_Number := 7;
   GC07_RC04.Hardware_U03.Speed1 := 500;
   GC07_RC04.Hardware_U03.RefSpeed := 1000;
   GC07_RC04.Hardware_U03.RD1_Motor_Number := 8;
   GC07_RC04.Hardware_U03.RD2_Motor_Number := 9;
   GC07_RC04.Hardware_U03.RD3_Motor_Number := 10;
   GC07_RC05.Hardware_U01.Speed1 := 500;
   GC07_RC05.Hardware_U01.RefSpeed := 1000;
   GC07_RC05.Hardware_U01.RD1_Motor_Number := 1;
   GC07_RC05.Hardware_U01.RD2_Motor_Number := 2;
   GC07_RC05.Hardware_U01.RD3_Motor_Number := 3;
   GC07_RC06.Hardware_U01.Speed1 := 500;
   GC07_RC06.Hardware_U01.RefSpeed := 1000;
   GC07_RC06.Hardware_U01.RD1_Motor_Number := 1;
   GC07_RC06.Hardware_U01.RD2_Motor_Number := 2;
   GC07_RC10.Hardware_U01.Speed1 := 500;
   GC07_RC10.Hardware_U01.RefSpeed := 1000;
   GC07_RC10.Hardware_U01.RD3_Motor_Number := 1;
   GC07_RC10.Hardware_U01.RD4_Motor_Number := 2;
   GC07_RC07.Hardware_U01.Speed1 := 500;
   GC07_RC07.Hardware_U01.RefSpeed := 1000;
   GC07_RC07.Hardware_U01.RD1_Motor_Number := 1;
   GC07_RC07.Hardware_U01.RD2_Motor_Number := 2;
   GC07_RC07.Hardware_U01.RD3_Motor_Number := 3;
   GC07_RC07.Hardware_U01.RD4_Motor_Number := 4;
   GC07_RC07.Hardware_U02.Speed1 := 500;
   GC07_RC07.Hardware_U02.RefSpeed := 1000;
   GC07_RC07.Hardware_U02.RD1_Motor_Number := 5;
   GC07_RC07.Hardware_U02.RD2_Motor_Number := 6;
   GC07_RC07.Hardware_U02.RD3_Motor_Number := 7;
   GC07_RC07.Hardware_U02.RD4_Motor_Number := 8;
   GC07_RC07.Hardware_U03.Speed1 := 500;
   GC07_RC07.Hardware_U03.RefSpeed := 1000;
   GC07_RC07.Hardware_U03.RD1_Motor_Number := 9;
   GC07_RC07.Hardware_U03.RD2_Motor_Number := 10;
   GC07_RC08.Hardware_U01.Speed1 := 500;
   GC07_RC08.Hardware_U01.RefSpeed := 1000;
   GC07_RC08.Hardware_U01.RD1_Motor_Number := 1;
   GC07_RC08.Hardware_U01.RD2_Motor_Number := 2;
   GC07_RC11.Hardware_U01.Speed1 := 500;
   GC07_RC11.Hardware_U01.RefSpeed := 1000;
   GC07_RC11.Hardware_U01.RD3_Motor_Number := 1;
   GC07_RC11.Hardware_U01.RD4_Motor_Number := 2;

END_DATA_BLOCK

FUNCTION_BLOCK "FB_Digital_Signal"
TITLE = FB_Digital_Signal
{ S7_Optimized_Access := 'TRUE' }
AUTHOR : 'Jay Liu'
VERSION : 0.1
//Filter digital signal with delay on and delay off
//
//[DESCRIPTION]
//Filter digital signal with delay on and delay off
//
//[BLOCK_INFO_HEADER]
//-------------------------------------------------------------------------------
// Title:            FB_Digital_Signal
// Comment/Function: Filter digital signal with delay on and delay off
// Library/Family:   APS
// Author:           Jay Liu
// Tested with:      ---
// Engineering:      TIA Portal V20
// Restrictions:     ---
// Requirements:     ---
//-------------------------------------------------------------------------------
// Change log table:
// Version  | Date       | Author                 | Description
//----------|------------|------------------------|------------------------------
// 01.00.00 | 2026-01-22 | Jay Liu                | First released version
   VAR_INPUT RETAIN
      i_Signal : Bool;   // Input signal
      i_CMD_Preset : Bool;   // Command for preset filterd signal
      i_CFG_Dealy_On : DInt;   // Delay on raising edge of signal
      i_CFG_Dealy_Off : DInt;   // Delay off trailing edge of signal
      i_Cycle_Count : DInt;   // Cycle step
   END_VAR

   VAR_OUTPUT RETAIN
      o_Signal_Filtered : Bool;   // Filtered Signal
      o_Signal_Raising_Edge : Bool;   // Raising edge of filterd signal
      o_Signal_Trailing_Edge : Bool;   // Trailing edge of filterd signal
   END_VAR

   VAR RETAIN
      s_Signal_Filtered : Bool;   // Filtered Signal
      s_Copy_Signal : Bool;   // Previous state of input signal
      s_Copy_Signal_Filtered : Bool;   // Previous state of filterd signal
      s_Count_Filter : DInt;   // Count of filter
   END_VAR


BEGIN
	// Monitor change event
	IF #i_Signal XOR #s_Signal_Filtered THEN
	    IF #i_Signal AND NOT #s_Copy_Signal THEN
	        #s_Count_Filter := #i_CFG_Dealy_On;
	    END_IF;

	    IF NOT #i_Signal AND #s_Copy_Signal THEN
	        #s_Count_Filter := #i_CFG_Dealy_Off;
	    END_IF;

	    IF #i_CMD_Preset THEN
	        #s_Count_Filter := 0;
	    END_IF;
	END_IF;

	// Timer
	IF #i_Signal XOR #s_Signal_Filtered THEN
	    #s_Count_Filter := #s_Count_Filter - #i_Cycle_Count;
	    IF #s_Count_Filter < 0 THEN
	        #s_Count_Filter := 0;
	    END_IF;
	END_IF;

	IF #s_Count_Filter <= 0 THEN
	    #s_Signal_Filtered := #i_Signal;
	END_IF;

	// Output
	#o_Signal_Filtered := #s_Signal_Filtered;
	#o_Signal_Raising_Edge := #s_Signal_Filtered AND NOT #s_Copy_Signal_Filtered;
	#o_Signal_Trailing_Edge := NOT #s_Signal_Filtered AND #s_Copy_Signal_Filtered;
	#s_Copy_Signal_Filtered := #s_Signal_Filtered;
	#s_Copy_Signal := #i_Signal;
END_FUNCTION_BLOCK

TYPE "UDT_S210_HW_Interface"
VERSION : 0.1
   STRUCT
      Input { S7_SetPoint := 'False'} : "UDT_S210_HW_Input";
      Output { S7_SetPoint := 'False'} : "UDT_S210_HW_Output";
   END_STRUCT;

END_TYPE

FUNCTION_BLOCK "FB_SWS_Array_Control"
{ S7_Optimized_Access := 'TRUE' }
VERSION : 0.1
   VAR_INPUT
      i_CMD_Roller_Run : Bool;
      i_CMD_Straight : Bool;
      i_CMD_Divert_Left : Bool;
      i_CMD_Divert_Right : Bool;
      i_CMD_Manual_Mode : Bool;
      i_CMD_Fixed_Straight : Bool;
      i_CMD_Fixed_Left : Bool;
      i_CMD_Fixed_Right : Bool;
      i_CMD_Fixed_Ratio : Bool;
      i_New_Item_Present : Bool;
      i_Cycle_Count : Int;
      i_Setting : "UDT_SWS_Divert_Setting";
      i_Servos_Status : Array[1..#C_ARRAY_COUNT] of "UDT_SWS_Servo_Status";
   END_VAR

   VAR_IN_OUT
      io_Global : "UDT_Global";
      io_Array_Command : Array[1..#C_ARRAY_COUNT] of Struct
         CMD_Straight : Bool;
         CMD_Left : Bool;
         CMD_Right : Bool;
      END_STRUCT;
      io_Roller_IO_Interface : "UDT_SWS_Roller_IO";
   END_VAR

   VAR
      s_CMD_Straight : Bool;
      s_CMD_Left : Bool;
      s_CMD_Right : Bool;
      s_Mode_Fixed_Ratio : Bool;
      s_Mode_Auto : Bool;
      s_Copy_CMD_Straight : Bool;
      s_Copy_CMD_Left : Bool;
      s_Copy_CMD_Right : Bool;
      s_Copy_Mode_Fixed_Ratio : Bool;
      s_Copy_Mode_Auto : Bool;
      s_Copy_New_Item_Present : Bool;
      s_OS_New_Item_Present : Bool;
      s_Cnt_Item_Straight : Int;
      s_Cnt_Item_Left : Int;
      s_Cnt_Item_Right : Int;
      s_Array_Control : Array[1..#C_ARRAY_COUNT] of Struct
         Delay_Time : Int;
         Count_Delay_Time : Int;
         Run_Dwn_Delay { S7_SetPoint := 'True'} : Bool;
      END_STRUCT;
   END_VAR

   VAR_TEMP
      t_Index : UInt;
      t_Announce_Downstream : Bool;
   END_VAR

   VAR CONSTANT
      C_ARRAY_COUNT : UInt := 9;
   END_VAR


BEGIN
	REGION Build Configuration
	    #s_Array_Control[1].Delay_Time := #i_Setting.Group2_Action_Delay;
	    #s_Array_Control[2].Delay_Time := #i_Setting.Group3_Action_Delay;
	    #s_Array_Control[3].Delay_Time := #i_Setting.Group4_Action_Delay;
	    #s_Array_Control[4].Delay_Time := #i_Setting.Group5_Action_Delay;
	    #s_Array_Control[5].Delay_Time := #i_Setting.Group6_Action_Delay;
	    #s_Array_Control[6].Delay_Time := #i_Setting.Group7_Action_Delay;
	    #s_Array_Control[7].Delay_Time := #i_Setting.Group8_Action_Delay;
	    #s_Array_Control[8].Delay_Time := #i_Setting.Group9_Action_Delay;
	END_REGION

	REGION Handle Command
	    #s_CMD_Straight := (#i_CMD_Straight AND NOT #i_CMD_Divert_Left AND NOT #i_CMD_Divert_Right AND NOT #i_CMD_Manual_Mode)
	    OR (#i_CMD_Fixed_Straight AND NOT #i_CMD_Fixed_Left AND NOT #i_CMD_Fixed_Right AND #i_CMD_Manual_Mode);

	    #s_CMD_Left := (NOT #i_CMD_Straight AND #i_CMD_Divert_Left AND NOT #i_CMD_Divert_Right AND NOT #i_CMD_Manual_Mode)
	    OR (NOT #i_CMD_Fixed_Straight AND #i_CMD_Fixed_Left AND NOT #i_CMD_Fixed_Right AND #i_CMD_Manual_Mode);

	    #s_CMD_Right := (NOT #i_CMD_Straight AND NOT #i_CMD_Divert_Left AND #i_CMD_Divert_Right AND NOT #i_CMD_Manual_Mode)
	    OR (NOT #i_CMD_Fixed_Straight AND NOT #i_CMD_Fixed_Left AND #i_CMD_Fixed_Right AND #i_CMD_Manual_Mode);

	    #s_Mode_Fixed_Ratio := #i_CMD_Fixed_Ratio AND #i_CMD_Manual_Mode;
	END_REGION

	REGION Fixed Ratio Mode
	    #s_OS_New_Item_Present := #i_New_Item_Present AND NOT #s_Copy_New_Item_Present;
	    IF #s_Mode_Fixed_Ratio THEN

	        IF #s_Cnt_Item_Straight <= 0 AND #s_Cnt_Item_Left <= 0 AND #s_Cnt_Item_Right <= 0 THEN
	            #s_Cnt_Item_Straight := #i_Setting.Fixed_Ratio_Staight;
	            #s_Cnt_Item_Left := #i_Setting.Fixed_Ratio_Left;
	            #s_Cnt_Item_Right := #i_Setting.Fixed_Ratio_Right;
	        END_IF;

	        IF #s_OS_New_Item_Present THEN
	            IF #s_Cnt_Item_Left > 0 THEN
	                #s_Array_Control[1].Run_Dwn_Delay := TRUE;
	                #io_Array_Command[1].CMD_Straight := FALSE;
	                #io_Array_Command[1].CMD_Left := TRUE;
	                #io_Array_Command[1].CMD_Right := FALSE;
	                #s_Array_Control[1].Count_Delay_Time := 0;
	                #s_Cnt_Item_Left -= 1;
	            ELSIF #s_Cnt_Item_Straight > 0 THEN
	                #s_Array_Control[1].Run_Dwn_Delay := TRUE;
	                #io_Array_Command[1].CMD_Straight := TRUE;
	                #io_Array_Command[1].CMD_Left := FALSE;
	                #io_Array_Command[1].CMD_Right := FALSE;
	                #s_Array_Control[1].Count_Delay_Time := 0;
	                #s_Cnt_Item_Straight -= 1;
	            ELSIF #s_Cnt_Item_Right > 0 THEN
	                #s_Array_Control[1].Run_Dwn_Delay := TRUE;
	                #io_Array_Command[1].CMD_Straight := FALSE;
	                #io_Array_Command[1].CMD_Left := FALSE;
	                #io_Array_Command[1].CMD_Right := TRUE;
	                #s_Array_Control[1].Count_Delay_Time := 0;
	                #s_Cnt_Item_Right -= 1;
	            END_IF;
	        END_IF;
	    END_IF;
	END_REGION

	REGION Divert Command
	    IF #s_CMD_Straight AND NOT #s_Copy_CMD_Straight THEN
	        #s_Array_Control[1].Run_Dwn_Delay := TRUE;
	        #io_Array_Command[1].CMD_Straight := TRUE;
	        #io_Array_Command[1].CMD_Left := FALSE;
	        #io_Array_Command[1].CMD_Right := FALSE;
	        #s_Array_Control[1].Count_Delay_Time := 0;
	    END_IF;

	    IF #s_CMD_Left AND NOT #s_Copy_CMD_Left THEN
	        #s_Array_Control[1].Run_Dwn_Delay := TRUE;
	        #io_Array_Command[1].CMD_Straight := FALSE;
	        #io_Array_Command[1].CMD_Left := TRUE;
	        #io_Array_Command[1].CMD_Right := FALSE;
	        #s_Array_Control[1].Count_Delay_Time := 0;
	    END_IF;

	    IF #s_CMD_Right AND NOT #s_Copy_CMD_Right THEN
	        #s_Array_Control[1].Run_Dwn_Delay := TRUE;
	        #io_Array_Command[1].CMD_Straight := FALSE;
	        #io_Array_Command[1].CMD_Left := FALSE;
	        #io_Array_Command[1].CMD_Right := TRUE;
	        #s_Array_Control[1].Count_Delay_Time := 0;
	    END_IF;
	END_REGION

	FOR #t_Index := 1 TO #C_ARRAY_COUNT DO
	    "FC_Delay_On_Accumulator"(i_CMD_Start    := #s_Array_Control[#t_Index].Run_Dwn_Delay,
	                              i_Enable_Dly   := #i_CMD_Roller_Run,
	                              i_CFG_Target   := #s_Array_Control[#t_Index].Delay_Time,
	                              i_Cycle_Count  := #i_Cycle_Count,
	                              o_Delay_Finish => #t_Announce_Downstream,
	                              io_Setpoint    := #s_Array_Control[#t_Index].Count_Delay_Time);

	    IF #t_Index < #C_ARRAY_COUNT AND #t_Announce_Downstream THEN
	        #s_Array_Control[#t_Index].Run_Dwn_Delay := FALSE;
	        #s_Array_Control[#t_Index + 1].Run_Dwn_Delay := TRUE;
	        #io_Array_Command[#t_Index + 1].CMD_Straight := #io_Array_Command[#t_Index].CMD_Straight;
	        #io_Array_Command[#t_Index + 1].CMD_Left := #io_Array_Command[#t_Index].CMD_Left;
	        #io_Array_Command[#t_Index + 1].CMD_Right := #io_Array_Command[#t_Index].CMD_Right;
	    END_IF;
	END_FOR;

	REGION Control Roller Speed
	    #io_Roller_IO_Interface.Output.Array1_Speed1 := #i_CMD_Roller_Run AND NOT #io_Array_Command[1].CMD_Left;
	    #io_Roller_IO_Interface.Output.Array1_Speed2 := #i_CMD_Roller_Run AND (#io_Array_Command[1].CMD_Left OR #io_Array_Command[1].CMD_Right);
	    #io_Roller_IO_Interface.Output.Array2_Speed1 := #i_CMD_Roller_Run AND NOT #io_Array_Command[2].CMD_Left;
	    #io_Roller_IO_Interface.Output.Array2_Speed2 := #i_CMD_Roller_Run AND (#io_Array_Command[2].CMD_Left OR #io_Array_Command[2].CMD_Right);
	    #io_Roller_IO_Interface.Output.Array3_Speed1 := #i_CMD_Roller_Run AND NOT #io_Array_Command[3].CMD_Left;
	    #io_Roller_IO_Interface.Output.Array3_Speed2 := #i_CMD_Roller_Run AND (#io_Array_Command[3].CMD_Left OR #io_Array_Command[3].CMD_Right);
	    #io_Roller_IO_Interface.Output.Array4_Speed1 := #i_CMD_Roller_Run AND NOT #io_Array_Command[4].CMD_Left;
	    #io_Roller_IO_Interface.Output.Array4_Speed2 := #i_CMD_Roller_Run AND (#io_Array_Command[4].CMD_Left OR #io_Array_Command[4].CMD_Right);
	    #io_Roller_IO_Interface.Output.Array5_Speed1 := #i_CMD_Roller_Run AND NOT #io_Array_Command[5].CMD_Left;
	    #io_Roller_IO_Interface.Output.Array5_Speed2 := #i_CMD_Roller_Run AND (#io_Array_Command[5].CMD_Left OR #io_Array_Command[5].CMD_Right);
	    #io_Roller_IO_Interface.Output.Array6_Speed1 := #i_CMD_Roller_Run AND NOT #io_Array_Command[6].CMD_Left;
	    #io_Roller_IO_Interface.Output.Array6_Speed2 := #i_CMD_Roller_Run AND (#io_Array_Command[6].CMD_Left OR #io_Array_Command[6].CMD_Right);
	    #io_Roller_IO_Interface.Output.Array7_Speed1 := #i_CMD_Roller_Run AND NOT #io_Array_Command[7].CMD_Left;
	    #io_Roller_IO_Interface.Output.Array7_Speed2 := #i_CMD_Roller_Run AND (#io_Array_Command[7].CMD_Left OR #io_Array_Command[7].CMD_Right);
	    #io_Roller_IO_Interface.Output.Array8_Speed1 := #i_CMD_Roller_Run AND NOT #io_Array_Command[8].CMD_Left;
	    #io_Roller_IO_Interface.Output.Array8_Speed2 := #i_CMD_Roller_Run AND (#io_Array_Command[8].CMD_Left OR #io_Array_Command[8].CMD_Right);
	    #io_Roller_IO_Interface.Output.Array9_Speed1 := #i_CMD_Roller_Run AND NOT #io_Array_Command[9].CMD_Left;
	    #io_Roller_IO_Interface.Output.Array9_Speed2 := #i_CMD_Roller_Run AND (#io_Array_Command[9].CMD_Left OR #io_Array_Command[9].CMD_Right);
	END_REGION

	REGION Storage Previous State
	    #s_Copy_CMD_Straight := #s_CMD_Straight;
	    #s_Copy_CMD_Left := #s_CMD_Left;
	    #s_Copy_CMD_Right := #s_CMD_Right;
	    #s_Copy_Mode_Fixed_Ratio := #s_Mode_Fixed_Ratio;
	    #s_Copy_Mode_Auto := #s_Mode_Auto;
	    #s_Copy_New_Item_Present := #i_New_Item_Present;
	END_REGION

END_FUNCTION_BLOCK

TYPE "UDT_Conv_S210_Command"
VERSION : 0.1
   STRUCT
      Man_Mode : Bool := false;   // Maintenance mode on
      Man_Clear : Bool := false;   // Maintenance - Clear data
      Man_Run : Bool := false;   // Maintenance - Run motor
      Man_DisableAxis : Bool;   // Maintenance - Disable axis
      Cmd_Reset_ESave : Bool := false;   // Command - Reset energy save
      Cmd_Bypass_Fault : Bool := false;   // Command - Bypass all fault
      Spare_0_6 : Bool := false;   // Spare_0_6
      Spare_0_7 : Bool := false;   // Spare_0_7
      Spare_1_0 : Bool := false;   // Spare_1_0
      Spare_1_1 : Bool := false;   // Spare_1_1
      Spare_1_2 : Bool := false;   // Spare_1_2
      Spare_1_3 : Bool := false;   // Spare_1_3
      Spare_1_4 : Bool := false;   // Spare_1_4
      Spare_1_5 : Bool := false;   // Spare_1_5
      Spare_1_6 : Bool := false;   // Spare_1_6
      Spare_1_7 : Bool := false;   // Spare_1_7
   END_STRUCT;

END_TYPE

FUNCTION_BLOCK "FB_HW_SWS_S210"
{ S7_Optimized_Access := 'TRUE' }
VERSION : 0.1
   VAR_INPUT
      i_Telegram_HW_ID : HW_SUBMODULE;
      i_Additional_HW_ID { ExternalAccessible := 'False'; ExternalVisible := 'False'; ExternalWritable := 'False'} : HW_SUBMODULE;
      i_IO_Available : Bool;
      i_Safety_OK : Bool := TRUE;
      i_CMD_Reset : Bool;
      i_CMD_Maintenance_Mode : Bool;
      i_CMD_Disable_Axis : Bool;
      i_CMD_Home : Bool;
      i_CMD_Jog_Left : Bool;
      i_CMD_Jog_Right : Bool;
      i_CMD_Save : Bool;
      i_CMD_Straight : Bool;
      i_CMD_Divert_Left : Bool;
      i_CMD_Divert_Right : Bool;
      i_HW_Setting : "UDT_SWS_Servo_Setting";
   END_VAR

   VAR_OUTPUT RETAIN
      o_Ready_To_Reset : Bool;
      o_ER_PN_Not_Present : Bool;
      o_ER_PN_Error : Bool;
      o_ST_Axis_Enabled : Bool;
      o_ST_Position_Reached : Bool;
      o_OL_Maintenance_Mode : Bool;
      o_ER_Motor_Fault : Bool;
      o_ER_Home_Position_Missing : Bool;
      o_ER_STO_Active : Bool;
      o_WN_Motor_Alarm : Bool;
      o_ST_Act_Position : Real;
      o_AlarmCode : Word;
      o_FaultCode : Word;
   END_VAR

   VAR_IN_OUT
      io_Global : "UDT_Global";
      io_S210_Interface : "UDT_S210_HW_Interface";
   END_VAR

   VAR
      s_FB_SINA_POS_TEL112 : "FB_SINA_POS_TEL112";
      s_FB_SINA_Save_Parameter : "FB_SINA_Save_Parameter";
   END_VAR
   VAR RETAIN
      s_SW_In { S7_SetPoint := 'False'} : "UDT_S210_SW_Input";
      s_SW_Out { S7_SetPoint := 'False'} : "UDT_S210_SW_Output";
      s_Actual_Value : Struct
         ZSW_S210_Bit08_Reserved : Bool;
         ZSW_S210_Bit09_Reserved : Bool;
         ZSW_S210_Bit10_Reserved : Bool;
         ZSW_S210_Bit11_Reserved : Bool;
         ZSW_S210_Bit12_Reserved : Bool;
         ZSW_S210_Bit13_Reserved : Bool;
         ZSW_S210_Bit14_Reserved : Bool;
         ZSW_S210_Bit15_Reserved : Bool;
         ZSW_S210_Bit00_DI0 : Bool;
         ZSW_S210_Bit01_DI1 : Bool;
         ZSW_S210_Bit02_DI2 : Bool;
         ZSW_S210_Bit03_DI3 : Bool;
         ZSW_S210_Bit04_DI4 : Bool;
         ZSW_S210_Bit05_Reserved : Bool;
         ZSW_S210_Bit06_Reserved : Bool;
         ZSW_S210_Bit07_Reserved : Bool;
         DCLinkVoltage : Int;
         ActualCurrent : Int;
         ActivePower : Int;
      END_STRUCT;
      s_Timer_Reset_Delay { S7_SetPoint := 'True'} : Int;
      s_Copy_CMD_Straight : Bool;
      s_Copy_CMD_Left : Bool;
      s_Copy_CMD_Right : Bool;
      s_Copy_CMD_Save : Bool;
   END_VAR

   VAR_TEMP
      t_GeoAddr {InstructionName := 'GEOADDR'; LibVersion := '1.0'} : GEOADDR;
      t_Ret_Val_Int : Int;   // Temp: Return Value Int
      t_Start_Address : Int;
      t_IO_Available : Bool;
      t_Actual_Telegram_HWID : HW_ANY;
   END_VAR

   VAR CONSTANT
      C_RESET_DELAY_TIME : Int := 200;
      C_MODE_ABSOLUTE_POSITION : Int := 2;
      C_MODE_SET_HOME_POSITION : Int := 5;
      C_MODE_JOG : Int := 7;
      C_MODE_ADJUST_ENCODER : Int := 9;
   END_VAR


BEGIN
	REGION NETOWRK: Initial
	    #o_Ready_To_Reset := FALSE;
	END_REGION

	REGION NETOWRK: Diagnose PN Status
	    #t_Ret_Val_Int := LOG2GEO(LADDR := #i_Telegram_HW_ID, GEOADDR := #t_GeoAddr);
	    IF #i_CMD_Reset OR NOT #i_IO_Available THEN
	        #o_ER_PN_Not_Present := FALSE;
	        #o_ER_PN_Error := FALSE;
	    END_IF;
	    IF #i_IO_Available AND (#t_Ret_Val_Int <> 0 OR "DB_Diagnostics".PNIO_System_100.Device_Not_Present[#t_GeoAddr.STATION]) THEN
	        #o_ER_PN_Not_Present := TRUE;
	    END_IF;
	    IF #i_IO_Available AND "DB_Diagnostics".PNIO_System_100.Device_Error[#t_GeoAddr.STATION] THEN
	        #o_ER_PN_Error := TRUE;
	    END_IF;
	    IF
	        #o_ER_PN_Not_Present AND NOT (#t_Ret_Val_Int <> 0 OR "DB_Diagnostics".PNIO_System_100.Device_Not_Present[#t_GeoAddr.STATION])
	        //OR (#o_ER_PN_Error AND NOT ""DB_Diagnostics"".PNIO_System_100.Device_Error[#t_GeoAddr.STATION])
	    THEN
	        #o_Ready_To_Reset := TRUE;
	    END_IF;
	    #t_IO_Available := #i_IO_Available AND NOT #o_ER_PN_Not_Present;
	END_REGION

	REGION NETWORK: Read IO
	    IF NOT #io_Global.PLC_Is_Simulated THEN
	        "FC_IFM_VFD_S210_In"(i_Telegram_HW_ID            := #i_Telegram_HW_ID,
	                             i_Additional_HW_ID          := #i_Additional_HW_ID,
	                             o_Telegram_Start_Address    => #t_Start_Address,
	                             o_ActualValue_Start_Address => #t_Start_Address,
	                             o_Data                      => #io_S210_Interface.Input);
	    END_IF;
	END_REGION

	REGION NETOWRK: Fixed Value
	    #s_SW_In.OverV := 100;
	END_REGION

	REGION NETOWRK: Reset Pulse
	    "FC_Delay_Off"(i_CMD_Start     := #i_CMD_Reset AND #t_IO_Available,
	                   i_CFG_Target    := #C_RESET_DELAY_TIME,
	                   i_Cycle_Count   := #io_Global.OB_Prev_Cycle_Time,
	                   o_Delay_Finish => #s_SW_In.AckError,
	                   io_Setpoint     := #s_Timer_Reset_Delay);
	END_REGION

	REGION NETOWRK: Axis Enable
	    #s_SW_In.Enbale := NOT #i_CMD_Disable_Axis AND #t_IO_Available AND #i_Safety_OK AND NOT #s_SW_Out.Lockout AND NOT #s_SW_Out.AxisError;
	END_REGION

	REGION NETOWRK: Auto Mode
	    IF NOT #i_CMD_Maintenance_Mode THEN
	        #s_SW_In.Mode := #C_MODE_ABSOLUTE_POSITION;
	        #s_SW_In.ConfigEPOS := 16#00000003;
	        #s_SW_In.CancelTraversing := TRUE;
	        #s_SW_In.IntermediateStop := TRUE;
	        IF #i_HW_Setting.Enable_Soft_Limit THEN
	            #s_SW_In.ConfigEPOS.%X2 := TRUE;
	        END_IF;
	        IF #i_HW_Setting.Enable_Hard_Limit THEN
	            #s_SW_In.ConfigEPOS.%X3 := TRUE;
	        END_IF;
	        IF #i_HW_Setting.Continuous_Action_Mode THEN
	            #s_SW_In.ConfigEPOS.%X8 := TRUE;
	        END_IF;
	        #s_SW_In.Velocity := INT_TO_REAL(LIMIT_INT(MN := 0, IN := #i_HW_Setting.Speed_Setpoint, MX := #i_HW_Setting.Max_Speed));
	        #s_SW_In.Acceleration := INT_TO_REAL(#i_HW_Setting.Acc_Setpoint);
	        #s_SW_In.Deceleration := INT_TO_REAL(#i_HW_Setting.Dec_Setpoint);

	        IF #i_CMD_Straight THEN
	            #s_SW_In.Position := 0.0;
	        ELSIF #i_CMD_Divert_Left THEN
	            #s_SW_In.Position := INT_TO_REAL(LIMIT_INT(MN := #i_HW_Setting.Max_Left_Position, IN := #i_HW_Setting.Left_Position_Setpoint, MX := 0));
	        ELSIF #i_CMD_Divert_Right THEN
	            #s_SW_In.Position := INT_TO_REAL(LIMIT_INT(MN := 0, IN := #i_HW_Setting.Right_Position_Setpoint, MX := #i_HW_Setting.Max_Right_Position));
	        END_IF;

	        #s_SW_In.ExecuteMode := FALSE;
	        IF
	            (#i_CMD_Straight AND NOT #s_Copy_CMD_Straight
	            AND NOT #i_CMD_Divert_Left
	            AND NOT #i_CMD_Divert_Right)
	            OR (#i_CMD_Divert_Left AND NOT #s_Copy_CMD_Left
	            AND NOT #i_CMD_Straight
	            AND NOT #i_CMD_Divert_Right)
	            OR (#i_CMD_Divert_Right AND NOT #s_Copy_CMD_Right
	            AND NOT #i_CMD_Straight
	            AND NOT #i_CMD_Divert_Left)
	        THEN
	            #s_SW_In.ExecuteMode := TRUE;
	        END_IF;
	    END_IF;
	END_REGION

	REGION NETOWRK: Maintenance Mode
	    IF #i_CMD_Maintenance_Mode THEN
	        #s_SW_In.ExecuteMode := FALSE;

	        REGION Home Mode
	            IF
	                #i_CMD_Home
	                AND NOT (#i_CMD_Jog_Left OR #i_CMD_Jog_Right)
	            THEN
	                #s_SW_In.Mode := #C_MODE_ADJUST_ENCODER;
	                #s_SW_In.ExecuteMode := TRUE;
	            END_IF;
	        END_REGION

	        REGION Jog Mode
	            IF
	                (#i_CMD_Jog_Left
	                XOR #i_CMD_Jog_Right)
	                AND NOT #i_CMD_Home
	            THEN
	                #s_SW_In.Mode := #C_MODE_JOG;
	                #s_SW_In.ConfigEPOS := 16#00000003;
	                #s_SW_In.CancelTraversing := TRUE;
	                #s_SW_In.IntermediateStop := TRUE;
	                #s_SW_In.Jog_Left := #i_CMD_Jog_Left;
	                #s_SW_In.Jog_Right := #i_CMD_Jog_Right;
	                #s_SW_In.Positive := FALSE;
	                #s_SW_In.Negative := FALSE;
	            ELSE
	                #s_SW_In.Jog_Left := FALSE;
	                #s_SW_In.Jog_Right := FALSE;
	            END_IF;
	        END_REGION

	        REGION Save Parameter
	            #s_FB_SINA_Save_Parameter(i_Trigger  := #i_CMD_Save AND NOT #s_Copy_CMD_Save AND NOT (#i_CMD_Jog_Left OR #i_CMD_Jog_Right) AND NOT #i_CMD_Home,
	                                      i_VFD_Type := 2,
	                                      i_HW_ID    := #i_Telegram_HW_ID);
	            #s_Copy_CMD_Save := #i_CMD_Save;
	        END_REGION
	    END_IF;
	END_REGION

	 REGION NETOWRK: Siemens Telegram 112
	    #s_SW_In.ConfigEPOS.%X1 := #i_Safety_OK;

